(* IEC 61131-3 sources: daoli-st-library/DL_Process (part 71) *)

(* ---- FB_DL_ScrewConveyorDoseSeq.st ---- *)
(*==============================================================================
 * 组件名称 (Component)  : FB_DL_ScrewConveyorDoseSeq
 * 所属子库 (Sublibrary) : DL_Process ｜ 版本 (Version) : 1.0.0 ｜ 2026-11-24
 * 兼容性   (Platform)   : CODESYS 3.5+ / TwinCAT 3 / 汇川 InoProShop / 施耐德 Machine Expert
 *                         仅依赖 IEC 61131-3 标准库（TON / R_TRIG / ABS / MAX），零厂商私有库
 * 功能描述 (Function)   : 螺旋给料计量批次序列：预检 → 喂料（按 fFlowKgh × dt 定周期积算，
 *                         达提前量停料）→ 停料稳定 tSettle → 称量结算（算误差百分比、批次 +1、
 *                         发 bBatchDone 单拍）→ 完成相（bStart 仍 TRUE 则自动进入下一批）。
 *                         **积算口径**：dt 由定周期采样节拍 tonDt（PT = 100ms 常数）生成，
 *                         积分步长 _fDtSec = TIME_TO_LREAL(DL_SCD_DT)，且入口做 dt > EPS 闸
 *                         （防 dt ≤ 0 / 非正步长导致积分反向或除零，R4）；非采样拍不积分。
 *                         **提前量**：停料阈值 _fStopThr := fTargetKg × (1 − fTolPct/100)，
 *                         使停料后的空中料流残量落进容差带；eWeigh 再按实际 fDosedKg 结算。
 *                         **bStart = FALSE 语义（R191 二选一，本件选「降级为安全值 + 置标志」）**：
 *                         bMotorRun 落 FALSE 并回 eIdle（螺旋不得冻结保持，冻结即过量给料）。
 * 接口     (Interface)  : 输入 bEnable / bStart / bReset（上升沿）/ fTargetKg / fFlowKgh /
 *                         tSettle / tTimeout / fTolPct / bMotorFb；
 *                         输出 bMotorRun / fDosedKg / fErrPct / nBatchCnt / bBatchDone（单拍）/
 *                         eState（E_DL_ScdPhase）/ eCause（E_DL_ScdCause）/ bError / bValid。
 * 状态迁移表 (State Transition Table)：
 *   ① eIdle → ePreCheck：bEnable 且 bStart 且组态闸通过且 fTargetKg > 0 且无锁存；
 *      拍 N 进入 / 本拍行为：清 fDosedKg、fErrPct、nBatchCnt、bMotorRun=FALSE / 拍 N+1 转出。
 *   ② ePreCheck → eFeeding：预检相单拍驻留（本拍清零 fDosedKg / fErrPct，保证连续批次每批独立）；
 *      拍 N 进入 / 本拍行为：置 bMotorRun=TRUE / 拍 N+1 转出至 eFeeding。
 *   ③ eFeeding → eSettle：fDosedKg ≥ _fStopThr 或 fDosedKg ≥ fTargetKg（达量，事件优先于超时，
 *      FB51-5）；拍 N 进入 / 本拍行为：bMotorRun=FALSE、清积分节拍 / 拍 N+1 转出至 eSettle。
 *   ④ eSettle → eWeigh：tonSettle.Q（停料稳定到时）；拍 N 进入 / 本拍行为：bMotorRun=FALSE /
 *      拍 N+1 转出至 eWeigh。
 *   ⑤ eWeigh → eDone：单拍结算；本拍行为：nBatchCnt+1、置 _bBatchDoneInt（统一出口映射，
 *      FB33-1）、按 |fErrPct| 与 fTolPct 发 eBatchDone / eOutOfTol（均信息级）/ 拍 N+1 转出。
 *   ⑥ eDone → ePreCheck：bStart 仍 TRUE（连续批次）；拍 N 进入 / 本拍行为：bMotorRun=FALSE /
 *      拍 N+1 转出至 ePreCheck。⑦ eDone → eIdle：bStart 落 FALSE（前置消失，R98 两条出口）。
 *   ⑧ eFeeding → eFault：fFlowKgh < 0（eBadFlow，即时）/ 流量为 0 持续 tTimeout（eNoFlow）/
 *      总超时 tTimeout（eTimeout）/ bMotorRun 与 bMotorFb 不一致达 3s（eMotorNoFb）/
 *      全相入参非有限（eNonFinite）。锁存后由段尾迁移闸迁相（R21）。
 *   ⑨ eFault → eIdle：bReset 上升沿（R_TRIG 判 .Q）且 bEnable = FALSE（R19 穷举出口）；
 *      拍 N 进入 / 本拍行为：清锁存、成因、bMotorRun=FALSE / 拍 N+1 转出至 eIdle。
 *   ⑩ ELSE（非法枚举值）→ eFault，成因 eIllegalState（R6 兜底）。
 * 边界     (Boundary)   : ① 五个 TON 与 R_TRIG 全在 CASE 外无条件调用（R7）；tonDt / tonTotal /
 *                            tonNoFlow / tonSettle / tonMotFb 的 IN 均含 NOT .Q 自复位项（R188）。
 *                         ② 积分步长闸：_fDtSec > DL_SCD_EPS 才积分（R4 防 dt ≤ 0）；
 *                            fTargetKg ≤ EPS 时不做百分比除法，fErrPct 置 0 哨兵（除零不可达）。
 *                         ③ 浮点比较一律容差或大小比较，禁 `=`/`<>`（R4）；零流量判据为
 *                            ABS(fFlowKgh) < DL_SCD_EPS。
 *                         ④ 非有限判据：fTargetKg / fFlowKgh / fTolPct 逐拍双判（x<>x 判 NaN，
 *                            (x−x)<>0 判 Inf）。
 *                         ⑤ 无数组、无下标，故无越界风险；nBatchCnt 为 UDINT 单调累加不溢出。
 *                         ⑥ 零全局耦合（无 GVL / VAR_EXTERNAL / %I / %Q，R1 / R2）。
 * 码表     (Codes)      : 本件不占用全局数字码位（R297 零码位范式）；出口为 BOOL + ENUM，
 *                         enum E_DL_ScdPhase / E_DL_ScdCause 归属本文件（全库唯一属主，R264）。
 *                         信息级（0..9）永不置 bError；故障级（10 起）赋值处与 _bFaultLatch 三行
 *                         成对（R45），锁存回放至 bReset 沿（FB33-1）。
 * 分工声明 (Scope)      : 失重式连续给料控制（喂料闭环）归 FB_DL_ChemDosingGrav / FB_DL_BatchDosingControl；
 *                         批次报表与追溯归 DL_Process 报表件；本件只做**单批"喂料—稳定—称量"时序
 *                         与流量积算**，不做喂料闭环整定，也不做螺旋电机保护。
 * 归属     (Ownership)  : E_DL_ScdPhase / E_DL_ScdCause 归属本文件（全库唯一定义，R264）。
 * 红线自检 (Redline)    : R1 ✓ 零 GVL ｜ R2 ✓ 零 %I/%Q ｜ R3 ✓ 纯 IEC ｜ R4 ✓ dt 闸 + 除零闸 +
 *                         非有限双判 + 容差比较 ｜ R5 ✓ 逐行同行双语注释 ｜ R6 ✓ 七态 ENUM +
 *                         CASE + ELSE ｜ R7 ✓ 全部 TON/R_TRIG 在 CASE 外 ｜ R8/R9 N/A（无 METHOD）
 *                         R10 ✓ 无构造式转换（TIME_TO_LREAL / 标准函数）｜ R14 ✓ 无 PROPERTY
 *                         R15 ✓ 无保留字撞名 ｜ R17 ✓ 无数组｜ R18 ✓ bReset 用 R_TRIG 判 .Q
 *                         R19 ✓ eFault 出口 = bReset 沿 + 撤使能 ｜ R20 ✓ 稳定/供料等待相带超时
 *                         R21 ✓ 锁存与迁相分离。
 * 修订历史 (Revision)   : 2026-11-24  v1.0.0  R79-B 首版
 * 验收向量 (Acceptance) :
 *   V1 fTargetKg=10.0、fFlowKgh=3600.0（=1 kg/s）、fTolPct=1.0、tSettle=T#2S、tTimeout=T#60S：
 *      bEnable=bStart=TRUE → ePreCheck → eFeeding（bMotorRun=TRUE）；fDosedKg 每 100ms 增 0.1kg，
 *      达 9.9kg（_fStopThr）→ eSettle；2s 后 eWeigh → fErrPct≈−1.0、nBatchCnt=1、
 *      bBatchDone 单拍 TRUE（次拍 FALSE）→ eDone。
 *   V2 续 V1，bStart 保持 TRUE → eDone → ePreCheck 自动进入第 2 批；bStart 落 FALSE → 回 eIdle，
 *      nBatchCnt 清零。
 *   V3 fTargetKg=0.0 → eState=eFault、eCause=eBadConfig、bError=TRUE、bMotorRun=FALSE；
 *      bReset 上升沿且 bEnable=FALSE → 回 eIdle、bError=FALSE。
 *   V4 fFlowKgh=0.0 持续 tTimeout=T#5S → eState=eFault、eCause=eNoFlow、bError=TRUE。
 *   V5 fFlowKgh=−5.0（负流量）→ 当拍 eState=eFault、eCause=eBadFlow、bMotorRun=FALSE。
 *   V6 bMotorRun=TRUE 而 bMotorFb 保持 FALSE 超 3s → eState=eFault、eCause=eMotorNoFb。
 *============================================================================*)

(*-----------------------------------------------------------------------------
 * 枚举: E_DL_ScdPhase（螺旋给料批次相位；eFault 为安全相，仅 bReset 沿迁出）
 *----------------------------------------------------------------------------*)
TYPE E_DL_ScdPhase :
(
    eIdle     := 0,    // 空闲：电机停，计数值清零 / Idle: motor stopped, counters cleared
    ePreCheck := 10,   // 预检相：单拍，置电机启动命令 / Pre-check: single scan, arm the motor command
    eFeeding  := 20,   // 喂料相：电机运行，按流量 × dt 积算 / Feeding: motor on, integrate flow times dt
    eSettle   := 30,   // 稳定相：停料后等空中料流落净 / Settle: motor off, waiting for the in-flight material
    eWeigh    := 40,   // 称量相：单拍结算误差与批次 / Weigh: single-scan settlement of error and batch count
    eDone     := 50,   // 完成相：本批完成，等下一批或退出 / Done: batch finished, waiting for the next one
    eFault    := 90    // 故障安全相：锁存成因，电机全停 / Fault safe phase: latched cause, motor stopped
);
END_TYPE

(*-----------------------------------------------------------------------------
 * 枚举: E_DL_ScdCause（成因码；信息级 = 0..9，故障级 = 10 起）
 *----------------------------------------------------------------------------*)
TYPE E_DL_ScdCause :
(
    eNone       := 0,   // 信息级：无事件 / Info: no event
    eBatchDone  := 1,   // 信息级：一批完成且误差在容差内 / Info: batch completed within tolerance
    eOutOfTol   := 2,   // 信息级：一批完成但误差超容差（记录，不锁存）/ Info: batch completed out of tolerance, recorded only
    eSettling   := 3,   // 信息级：进入停料稳定相 / Info: entering the settle phase
    eBadConfig  := 10,  // 故障级：目标重量 / 容差 / 时间参数越域 / Fault: target, tolerance or time parameter out of domain
    eNonFinite  := 11,  // 故障级：入参非有限 / Fault: non-finite input
    eBadFlow    := 12,  // 故障级：流量为负 / Fault: negative flow
    eNoFlow     := 13,  // 故障级：流量为零持续超时（供料中断）/ Fault: zero flow persisted beyond the timeout
    eTimeout    := 14,  // 故障级：喂料总超时 / Fault: total feeding timeout
    eMotorNoFb  := 15,  // 故障级：电机命令与反馈不一致超 3s / Fault: motor command and feedback mismatch beyond 3 s
    eIllegalState := 16 // 故障级：非法状态枚举值 / Fault: illegal state enum value
);
END_TYPE

FUNCTION_BLOCK FB_DL_ScrewConveyorDoseSeq
VAR_INPUT
    bEnable    : BOOL := FALSE;        // 使能：FALSE 停电机并回 eIdle / Enable, FALSE stops the motor and returns to idle
    bStart     : BOOL := FALSE;        // 启动（电平）：FALSE 本批中止并回 eIdle / Start level, FALSE aborts the batch
    bReset     : BOOL := FALSE;        // 复位（上升沿，需同时 bEnable=FALSE）/ Reset rising edge, requires bEnable FALSE
    fTargetKg  : LREAL := 0.0;         // 批次目标重量，域 > 0 [kg] / Batch target weight, domain > 0
    fFlowKgh   : LREAL := 0.0;         // 当前给料流量（瞬时，来自流量计）[kg/h] / Instantaneous feed flow from the flow meter
    tSettle    : TIME := T#2S;         // 停料后稳定延时，域 0..1h [s] / Settle delay after the motor stops, domain 0..1h
    tTimeout   : TIME := T#60S;        // 喂料总超时，域 ≥ 100ms [s] / Total feeding timeout, domain >= 100ms
    fTolPct    : LREAL := 1.0;         // 允许误差，域 (0,100) [%] / Allowed error in percent, domain (0,100)
    bMotorFb   : BOOL := FALSE;        // 螺旋电机运行反馈（TRUE = 在转）[-] / Screw motor running feedback
END_VAR
VAR_OUTPUT
    bMotorRun  : BOOL;                 // 螺旋电机启动命令（电平）[-] / Screw motor run command, level
    fDosedKg   : LREAL := 0.0;         // 本批累计给料量 [kg] / Accumulated dose of this batch
    fErrPct    : LREAL := 0.0;         // 本批误差百分比（正 = 超量）[%] / Batch error percentage, positive means over-dose
    nBatchCnt  : UDINT := 0;           // 已完成批次数 [批] / Completed batch counter
    bBatchDone : BOOL;                 // 批次完成单拍脉冲（段 1 预置，统一出口映射）[-] / Single-scan batch-done pulse
    eState     : E_DL_ScdPhase;        // 状态出口（段尾单点映射）[-] / State outlet mapped at the tail
    eCause     : E_DL_ScdCause;        // 成因码出口（故障期锁存回放）[-] / Cause code outlet
    bError     : BOOL;                 // 故障锁存标志 [-] / Fault latch flag
    bValid     : BOOL;                 // 序列有效回执（喂料/稳定相且无锁存）[-] / Sequence validity receipt
END_VAR
VAR
    _eState      : E_DL_ScdPhase := E_DL_ScdPhase.eIdle;   // 内部相位（CASE 唯一写入目标）[-] / Internal phase
    _bFaultLatch : BOOL := FALSE;                          // 故障锁存位（仅 bReset 沿清除）[-] / Fault latch bit
    _eCauseLatch : E_DL_ScdCause := E_DL_ScdCause.eNone;    // 锁存成因码（FB33-1 锁存回放）[-] / Latched cause code
    _eCauseTmp   : E_DL_ScdCause := E_DL_ScdCause.eNone;    // 本拍首因中间量（段 8 组态闸用）[-] / First cause of this scan
    _bCfgOk      : BOOL := TRUE;                           // 组态与入参闸通过标志 [-] / Configuration gate flag
    _bResetPulse : BOOL := FALSE;                          // bReset 上升沿快照（R18）[-] / bReset rising-edge snapshot
    _bBatchDoneInt : BOOL := FALSE;                        // 批次完成内部单拍位（统一出口映射）[-] / Internal single-scan batch-done bit
    _fDtSec      : LREAL := 0.0;                           // 积分步长：[s] / Integration step in seconds
    _bDtOk       : BOOL := FALSE;                          // 积分步长有效性（dt > EPS）[-] / Integration step validity
    _fStopThr    : LREAL := 0.0;                           // 停料阈值 = 目标 × (1 − 容差%) [kg] / Stop threshold of the feed
    _fStepKg     : LREAL := 0.0;                           // 本采样拍积算增量 [kg] / Dose increment of this sampling scan
    _fErrCalc    : LREAL := 0.0;                           // 误差百分比中间量 [%] / Error percentage intermediate
    _bMotMismatch : BOOL := FALSE;                         // 电机命令与反馈不一致标志 [-] / Motor command and feedback mismatch
    _bMotRunPrev  : BOOL := FALSE;                         // 上一拍电机命令快照（段 4 不一致判据用，一拍延迟）/ Motor command snapshot of the last scan
    rtReset      : R_TRIG;                                 // bReset 边沿实例（段 4 无条件调用，R18）/ bReset edge instance called unconditionally
    tonDt        : TON;                                    // 定周期采样节拍（段 4 无条件调用）/ Fixed-period sampling tick
    tonTotal     : TON;                                    // 喂料总超时（段 4 无条件调用）/ Total feeding timeout
    tonNoFlow    : TON;                                    // 零流量持续判（段 4 无条件调用）/ Zero-flow persistence timer
    tonSettle    : TON;                                    // 停料稳定延时（段 4 无条件调用）/ Settle delay timer
    tonMotFb     : TON;                                    // 电机反馈不一致持续判（段 4 无条件调用）/ Motor feedback mismatch timer
END_VAR
VAR CONSTANT
    DL_SCD_ZERO      : LREAL := 0.0;            // 浮点零基准 [-] / Float zero base
    DL_SCD_ONE       : LREAL := 1.0;            // 浮点一基准 [-] / Float one base
    DL_SCD_HUNDRED   : LREAL := 100.0;          // 百分比基数 [%] / Percent base
    DL_SCD_SEC_HOUR  : LREAL := 3600.0;         // 每小时秒数（kg/h → kg）[s/h] / Seconds per hour converting kg/h to kg
    DL_SCD_EPS       : LREAL := 1.0E-6;         // 浮点同值/正步长容差 [-] / Float equality and positive-step tolerance
    DL_SCD_DT        : TIME := T#100MS;         // 采样节拍（积分步长来源）[s] / Sampling tick, the integration step source
    DL_SCD_FB_WIN    : TIME := T#3S;            // 电机反馈不一致持续窗 [s] / Motor feedback mismatch window
    DL_SCD_T_MIN     : TIME := T#100MS;         // 超时参数下限 [s] / Lower bound of the timeout parameters
    DL_SCD_T_MAX     : TIME := T#1H;            // 稳定/超时参数上限 [s] / Upper bound of the settle and timeout parameters
    DL_SCD_BATCH_INC : UDINT := 1;              // 批次计数步长（UDINT 显式常量）[批] / Batch counter increment
END_VAR

(* —— 段 1：单拍位与动作出口预置（不清锁存 / 累加量，FB32-1） —— *)
bBatchDone     := FALSE;                               // 单拍批次沿每拍预清 / Single-scan batch edge preset FALSE every scan
bMotorRun      := FALSE;                               // 电机命令预置（安全侧：默认不动作）/ Motor command preset, safe side
_bBatchDoneInt := FALSE;                               // 内部单拍位预清 / Internal single-scan bit preset
_bCfgOk        := TRUE;                                // 组态闸标志复位 / Configuration flag reset
_eCauseTmp     := E_DL_ScdCause.eNone;                  // 当拍首因复位 / Scan cause reset

(* —— 段 2：步长与阈值换算（浮点域闸前置） —— *)
_fDtSec   := TIME_TO_LREAL(DL_SCD_DT);                 // 采样节拍换算为秒（标准转换，R10）/ Sampling tick converted to seconds
IF _fDtSec > DL_SCD_EPS THEN
    _bDtOk := TRUE;                                    // 步长为正：允许积分 / Positive step: integration allowed
ELSE
    _bDtOk := FALSE;                                   // 步长非正：拒绝积分（R4 防 dt <= 0）/ Non-positive step: integration refused
END_IF
_fStopThr := DL_SCD_ZERO;                              // 停料阈值预置零 / Stop threshold preset
_fErrCalc := DL_SCD_ZERO;                               // 误差中间量预置零 / Error intermediate preset

(* —— 段 3：组态与入参域闸（R272 全量枚举浮点与时间引脚） —— *)
IF (fTargetKg <> fTargetKg) OR ((fTargetKg - fTargetKg) <> DL_SCD_ZERO)
    OR (fFlowKgh <> fFlowKgh) OR ((fFlowKgh - fFlowKgh) <> DL_SCD_ZERO)
    OR (fTolPct <> fTolPct) OR ((fTolPct - fTolPct) <> DL_SCD_ZERO) THEN
    _bCfgOk    := FALSE;                               // 入参非有限 / Non-finite input
    _eCauseTmp := E_DL_ScdCause.eNonFinite;            // 故障级：非有限入参 / Fault: non-finite input
END_IF
IF _bCfgOk THEN
    IF fTargetKg <= DL_SCD_EPS THEN
        _bCfgOk    := FALSE;                           // 目标重量非正 / Target weight not positive
        _eCauseTmp := E_DL_ScdCause.eBadConfig;        // 故障级：组态非法 / Fault: bad configuration
    ELSIF (fTolPct <= DL_SCD_EPS) OR (fTolPct >= DL_SCD_HUNDRED) THEN
        _bCfgOk    := FALSE;                           // 容差越域（0,100）/ Tolerance out of domain
        _eCauseTmp := E_DL_ScdCause.eBadConfig;        // 故障级：组态非法 / Fault: bad configuration
    ELSIF (tTimeout < DL_SCD_T_MIN) OR (tTimeout > DL_SCD_T_MAX) THEN
        _bCfgOk    := FALSE;                           // 超时参数越域 / Timeout out of domain
        _eCauseTmp := E_DL_ScdCause.eBadConfig;        // 故障级：组态非法 / Fault: bad configuration
    ELSIF tSettle > DL_SCD_T_MAX THEN
        _bCfgOk    := FALSE;                           // 稳定延时越上限 / Settle delay above the upper bound
        _eCauseTmp := E_DL_ScdCause.eBadConfig;        // 故障级：组态非法 / Fault: bad configuration
    ELSIF fFlowKgh < DL_SCD_ZERO THEN
        _bCfgOk    := FALSE;                           // 流量为负（传感器或工艺异常）/ Negative flow from the meter or process
        _eCauseTmp := E_DL_ScdCause.eBadFlow;          // 故障级：负流量 / Fault: negative flow
    END_IF
END_IF
IF _bCfgOk THEN
    (* 停料阈值 = 目标 × (1 − 容差%/100)；除数 100 为常量，除零结构性不可达 *)
    _fStopThr := fTargetKg * (DL_SCD_ONE - (fTolPct / DL_SCD_HUNDRED));
    IF _fStopThr <= DL_SCD_ZERO THEN
        _fStopThr := DL_SCD_ZERO;                      // 阈值负值兜底归零 / Clamp a negative threshold to zero
    END_IF
END_IF

(* —— 段 4：边沿与定时器（CASE 外无条件调用，R7；IN 均含 NOT .Q 自复位，R188） —— *)
rtReset(CLK := bReset);                                // bReset 边沿无条件刷新（R18）/ bReset edge refreshed unconditionally
_bResetPulse := rtReset.Q;                             // 边沿快照 / Edge snapshot
tonDt(IN := (_eState = E_DL_ScdPhase.eFeeding) AND (NOT tonDt.Q) AND (NOT _bFaultLatch),
      PT := DL_SCD_DT);                                // 喂料相定周期积分节拍 / Fixed-period integration tick while feeding
tonTotal(IN := (_eState = E_DL_ScdPhase.eFeeding) AND (NOT tonTotal.Q) AND (NOT _bFaultLatch),
         PT := tTimeout);                              // 喂料总超时 / Total feeding timeout
tonNoFlow(IN := (_eState = E_DL_ScdPhase.eFeeding) AND (ABS(fFlowKgh) < DL_SCD_EPS)
               AND (NOT tonNoFlow.Q) AND (NOT _bFaultLatch),
          PT := tTimeout);                             // 零流量持续判（供料中断）/ Zero-flow persistence check
tonSettle(IN := (_eState = E_DL_ScdPhase.eSettle) AND (NOT tonSettle.Q) AND (NOT _bFaultLatch),
          PT := tSettle);                              // 停料稳定延时 / Settle delay
_bMotMismatch := (_bMotRunPrev AND (NOT bMotorFb)) OR ((NOT _bMotRunPrev) AND bMotorFb);   // 命令与反馈不一致（用上一拍命令快照）/ Command and feedback mismatch using the last-scan command
tonMotFb(IN := _bMotMismatch AND (_eState = E_DL_ScdPhase.eFeeding)
              AND (NOT tonMotFb.Q) AND (NOT _bFaultLatch),
         PT := DL_SCD_FB_WIN);                         // 仅喂料相监视反馈一致性 / Feedback consistency monitored while feeding only

(* —— 段 5：误差百分比刷新（除零闸：目标重量非正时置零哨兵，R4） —— *)
IF fTargetKg > DL_SCD_EPS THEN
    _fErrCalc := ((fDosedKg - fTargetKg) / fTargetKg) * DL_SCD_HUNDRED;   // 误差百分比 / Error percentage
    fErrPct   := _fErrCalc;                                               // 误差出口 / Error outlet
ELSE
    fErrPct := DL_SCD_ZERO;                                               // 目标非正：置零哨兵（除零不可达）/ Zero sentinel, division unreachable
END_IF

(* —— 段 6：状态机主体（唯一相位写入点；故障只置锁存，迁相由段 8 统一执行） —— *)
CASE _eState OF
    E_DL_ScdPhase.eIdle :
        bMotorRun := FALSE;                            // 空闲：电机不动作 / Idle: motor idle
        fDosedKg  := DL_SCD_ZERO;                      // 累计量清零 / Dose counter cleared
        fErrPct   := DL_SCD_ZERO;                      // 误差清零 / Error cleared
        nBatchCnt := 0;                                // 批次计数清零 / Batch counter cleared
        IF bEnable AND bStart AND _bCfgOk AND (fTargetKg > DL_SCD_EPS) AND (NOT _bFaultLatch) THEN
            eCause  := E_DL_ScdCause.eNone;            // 信息级：无事件 / Info: no event
            _eState := E_DL_ScdPhase.ePreCheck;        // 迁移①：进入预检相 / Move to pre-check
        END_IF

    E_DL_ScdPhase.ePreCheck :
        IF (NOT bEnable) OR (NOT bStart) THEN
            bMotorRun := FALSE;                        // 失能：电机停 / Disabled: motor stopped
            eCause    := E_DL_ScdCause.eNone;          // 信息级：无事件 / Info: no event
            _eState   := E_DL_ScdPhase.eIdle;          // 回空闲相 / Back to idle
        ELSE
            fDosedKg  := DL_SCD_ZERO;                  // 每批起点：累计量清零 / Batch start: dose counter cleared
            fErrPct   := DL_SCD_ZERO;                  // 每批起点：误差清零 / Batch start: error cleared
            bMotorRun := TRUE;                         // 迁移②：预检通过，启动螺旋 / Pre-check passed: start the screw
            eCause    := E_DL_ScdCause.eNone;          // 信息级：无事件 / Info: no event
            _eState   := E_DL_ScdPhase.eFeeding;       // 进入喂料相 / Move to feeding
        END_IF

    E_DL_ScdPhase.eFeeding :
        bMotorRun := TRUE;                             // 喂料相电机保持运行 / Motor stays on while feeding
        IF (NOT bEnable) OR (NOT bStart) THEN
            bMotorRun := FALSE;                        // 失能：电机停 / Disabled: motor stopped
            eCause    := E_DL_ScdCause.eNone;          // 信息级：无事件 / Info: no event
            _eState   := E_DL_ScdPhase.eIdle;          // 回空闲相 / Back to idle
        ELSE
            (* 定周期积算：只有节拍拍且步长为正才积分（R4） *)
            IF tonDt.Q AND _bDtOk THEN
                _fStepKg  := (fFlowKgh * _fDtSec) / DL_SCD_SEC_HOUR;   // 增量 = 流量 × dt / 3600 [kg]
                fDosedKg  := fDosedKg + _fStepKg;                      // 累计给料量 / Accumulate the dose
            END_IF
            IF fFlowKgh < DL_SCD_ZERO THEN
                IF NOT _bFaultLatch THEN
                    _eCauseLatch := E_DL_ScdCause.eBadFlow;            // 故障级：负流量 / Fault: negative flow
                    _bFaultLatch := TRUE;                              // 置故障锁存（迁相由段 8，R21）/ Latch the fault
                END_IF
            ELSIF tonNoFlow.Q THEN
                IF NOT _bFaultLatch THEN
                    _eCauseLatch := E_DL_ScdCause.eNoFlow;             // 故障级：供料中断 / Fault: feed interrupted
                    _bFaultLatch := TRUE;                              // 置故障锁存 / Latch the fault
                END_IF
            ELSIF tonTotal.Q THEN
                IF NOT _bFaultLatch THEN
                    _eCauseLatch := E_DL_ScdCause.eTimeout;            // 故障级：喂料总超时 / Fault: total feeding timeout
                    _bFaultLatch := TRUE;                              // 置故障锁存 / Latch the fault
                END_IF
            ELSIF tonMotFb.Q THEN
                IF NOT _bFaultLatch THEN
                    _eCauseLatch := E_DL_ScdCause.eMotorNoFb;          // 故障级：电机反馈不一致 / Fault: motor feedback mismatch
                    _bFaultLatch := TRUE;                              // 置故障锁存 / Latch the fault
                END_IF
            ELSIF (fDosedKg >= _fStopThr) OR (fDosedKg >= fTargetKg) THEN
                bMotorRun := FALSE;                                    // 迁移③：达提前量，停料 / Reached the threshold: stop the feed
                eCause    := E_DL_ScdCause.eSettling;                  // 信息级：进入稳定相 / Info: entering settle
                _eState   := E_DL_ScdPhase.eSettle;                    // 进入稳定相 / Move to settle
            END_IF
        END_IF

    E_DL_ScdPhase.eSettle :
        bMotorRun := FALSE;                            // 稳定相电机保持停止 / Motor stays off while settling
        IF (NOT bEnable) OR (NOT bStart) THEN
            eCause  := E_DL_ScdCause.eNone;            // 信息级：无事件 / Info: no event
            _eState := E_DL_ScdPhase.eIdle;            // 回空闲相 / Back to idle
        ELSIF tonSettle.Q THEN
            eCause  := E_DL_ScdCause.eNone;            // 信息级：无事件 / Info: no event
            _eState := E_DL_ScdPhase.eWeigh;           // 迁移④：稳定到时进入称量相 / Settle elapsed: move to weigh
        END_IF

    E_DL_ScdPhase.eWeigh :
        bMotorRun      := FALSE;                       // 称量相电机停止 / Motor off during settlement
        nBatchCnt      := nBatchCnt + DL_SCD_BATCH_INC; // 迁移⑤：批次计数 +1 / Increment the batch counter
        _bBatchDoneInt := TRUE;                        // 批次完成内部单拍位置位 / Internal single-scan batch bit
        IF ABS(fErrPct) > fTolPct THEN
            eCause := E_DL_ScdCause.eOutOfTol;         // 信息级：误差超容差（记录，不锁存）/ Info: out of tolerance, recorded only
        ELSE
            eCause := E_DL_ScdCause.eBatchDone;        // 信息级：批次合格完成 / Info: batch completed within tolerance
        END_IF
        _eState := E_DL_ScdPhase.eDone;                // 进入完成相 / Move to done

    E_DL_ScdPhase.eDone :
        bMotorRun := FALSE;                            // 完成相电机停止 / Motor off in the done phase
        IF NOT bStart THEN
            eCause  := E_DL_ScdCause.eNone;            // 信息级：无事件 / Info: no event
            _eState := E_DL_ScdPhase.eIdle;            // 迁移⑦：前置消失回空闲 / Start gone: back to idle
        ELSIF NOT bEnable THEN
            eCause  := E_DL_ScdCause.eNone;            // 信息级：无事件 / Info: no event
            _eState := E_DL_ScdPhase.eIdle;            // 失能回空闲 / Disabled: back to idle
        ELSIF bStart AND bEnable THEN
            eCause  := E_DL_ScdCause.eNone;            // 信息级：无事件 / Info: no event
            _eState := E_DL_ScdPhase.ePreCheck;        // 迁移⑥：连续批次 / Continuous batches
        END_IF

    E_DL_ScdPhase.eFault :
        bMotorRun := FALSE;                            // 故障相：电机全停（安全侧）/ Fault phase: motor stopped
        IF _bResetPulse AND (NOT bEnable) THEN
            _bFaultLatch := FALSE;                     // 迁移⑨：清故障锁存 / Clear the fault latch
            _eCauseLatch := E_DL_ScdCause.eNone;       // 清锁存成因 / Clear the latched cause
            eCause       := E_DL_ScdCause.eNone;       // 出口同步归零 / Outlet follows
            fDosedKg     := DL_SCD_ZERO;               // 累计量清零 / Dose counter cleared
            fErrPct      := DL_SCD_ZERO;               // 误差清零 / Error cleared
            _eState      := E_DL_ScdPhase.eIdle;       // 回空闲相 / Back to idle
        END_IF

ELSE
    (* 迁移⑩：非法枚举兜底（R6） *)
    IF NOT _bFaultLatch THEN
        _eCauseLatch := E_DL_ScdCause.eIllegalState;   // 故障级：非法状态 / Fault: illegal state
        _bFaultLatch := TRUE;                          // 置故障锁存 / Latch the fault
    END_IF
END_CASE

(* —— 段 7：组态闸失败处理（锁存与迁相分离，R21） —— *)
IF (NOT _bCfgOk) AND (NOT _bFaultLatch) THEN
    _eCauseLatch := _eCauseTmp;                        // 锁存首因（组态闸）/ Latch the configuration cause
    _bFaultLatch := TRUE;                              // 置故障锁存 / Latch the fault
END_IF

(* —— 段 8：段尾故障迁移闸 + 故障相动作全撤（FB50-1④） —— *)
IF _bFaultLatch AND (_eState <> E_DL_ScdPhase.eFault) THEN
    _eState := E_DL_ScdPhase.eFault;                   // 锁存即迁相 / Latch forces the fault phase
END_IF
IF _eState = E_DL_ScdPhase.eFault THEN
    bMotorRun := FALSE;                                // 故障相动作全撤（含同拍迁入）/ Motor withdrawn in fault
END_IF

(* —— 段 9：统一出口（状态映射 + 单拍位映射 + 锁存回放） —— *)
eState     := _eState;                                 // 相位映射 / Phase mapping
bBatchDone := _bBatchDoneInt;                          // 单拍批次沿统一映射（FB33-1 两段式）/ Single-scan batch edge mapped here
bError     := _bFaultLatch;                            // 故障标志取锁存位 / Fault flag from the latch
IF _bFaultLatch THEN
    eCause := _eCauseLatch;                            // 故障期回放锁存码（FB33-1）/ Replay the latched code
END_IF
bValid := ((_eState = E_DL_ScdPhase.eFeeding) OR (_eState = E_DL_ScdPhase.eSettle))
          AND (NOT _bFaultLatch);                      // 喂料/稳定相且无锁存时有效 / Valid while feeding or settling without a latch
_bMotRunPrev := bMotorRun;                             // 电机命令快照更新（唯一写入点，段 4 用）/ Motor command snapshot, single write point
END_FUNCTION_BLOCK

(* ---- FB_DL_SipLineSterilSeq.st ---- *)
(*
    FB_DL_SipLineSterilSeq —— 管路 SIP 蒸汽灭菌顺控（排凝 → 升温 → 保温窗 → 冷却 → 放行）
    ------------------------------------------------------------------
    组件名称  : FB_DL_SipLineSterilSeq
    分类      : DL_Process / Sterilization
    前缀      : FB_DL_
    版本      : 1.0.0
    溯源      : 借鉴组织 —— T2-2 LBP 基础工艺（矩阵行 163）：仅借鉴
                「命令 → 监视 → 判定」三段分层骨架的公开语义；次源 T2-8
                ISA-88 相语义公开条款（相 / 状态命名惯例）；clean-room
                声明 —— 保温窗断点重计与温度判据 100% 自有，零代码行复制；
                SIP 121 ℃ 最低承诺属公开工程惯例条款（下界 100 ℃ 为本件
                组态锁存闸，可调）。
    平台      : 纯 IEC 61131-3（ENUM + CASE + TON / R_TRIG + TIME 算术），
                CODESYS 3.5 / TwinCAT 3 / InoProShop / Machine Expert 通用
    作者      : 道莅代码库 · PLC编程专家（R72 构建轮 · 批 4 · 序号 12）
    ------------------------------------------------------------------
    功能说明  : 管路蒸汽 SIP（Sterilize-In-Place）连续工艺段顺控：
                eIdle →（bEn ∧ 组态闸）eDrain（排凝，bDrainDone 反馈或
                tDrainTimeout 超时）→ eHeatUp（开蒸汽升温，fTempC 达
                fHoldTempSet 迁入）→ eHold（保温窗 TON 计时）→ eCooldown
                （关蒸汽，温度回落确认）→ eDone（bSterilized 放行保持）→
                eIdle（批界）。
                安全核心口径：
                ① fTempC 非有限（探头断线）→ **故障锁存 + 双输出立即关断**
                   ——温度状态不明不得放行，宁可重灭菌；
                ② 保温窗断点重计（SIP 无菌保证不容断点续计）：eHold 相内
                   fTempC 跌破 fHoldTempSet（每拍取本拍实时值，R42 本拍
                   复验口径）→ 计时中止回 eHeatUp + 扰动计数 +1，恢复后
                   TON 从零重计——断点续计等于伪造无菌时长，写死禁用；
                ③ fHoldTempSet 越承诺段（< 100 ℃）→ 组态锁存（SIP 公开
                   最低承诺 121 ℃ 工程惯例，下界闸定 100 ℃ 并留调参会空间
                   ——承诺下界以常量声明，单探头承诺段声明见边界八）；
                ④ 失能 → 双输出（bDrainCmd / bSteamCmd）清零 + bSterilized
                   撤销 + 状态回 eIdle（停机相输出清零，R57）；故障锁存保留，
                   复位沿解除；
                ⑤ 迁入 eHold 相与每拍判温均取本拍实时值（迁入拍即计时使能，
                   无跨拍陈旧判据）。
                冷却放行口径：eCooldown 以 fTempC < fHoldTempSet 确认回落
                （防高温放行烫尾），回落即 eDone；bSterilized 为**保持型**
                放行位（批界 = bEn 撤除或复位沿时清除）。
    错误码    : 16#0005_0640 工艺温度非有限（探头断线 / ADC 故障），双输出
                            立即关断，锁存至复位沿 —— 故障级
                16#0005_0641 排凝超时（eDrain 驻留超 tDrainTimeout），锁存
                            至复位沿 —— 故障级
                16#0005_0642 保温设定越承诺段（fHoldTempSet < 100 ℃ 或非
                            有限），锁存至复位沿 —— 故障级
                16#0005_0643 保温窗 / 排凝超时组态非正（tHoldTime /
                            tDrainTimeout <= 0），锁存至复位沿 —— 故障级
                加码反证句（R90）：0640 由「双输出关断 + eHealth 语义温度
                断线」唯一观测；0641 / 0642 / 0643 成因互斥且调用方可自证
                （反馈时序 / 组态表），输出组合（同为 eFault + bError）不可
                互换还原成因，维修动作各异，故各立一码；保温跌破扰动以
                uDisturbCount 专位观测（R90 不加码：扰动事件已有独立可观
                测出口，不重复发码）。
    码位总账  : 16#0005_0640 用 ｜ 16#0005_0641 用 ｜ 16#0005_0642 用 ｜
                16#0005_0643 用
                （0630 / 0631 已由 FB_DL_RejectBlowCtrl 占用，本件不占）
    边界与披露: 一 双 TON（tonDrain / tonHold）与 R_TRIG（rtReset）每拍
                   **无条件调用**（规则 ⑦），IN 为显式条件变量（R145 相驻留
                   口径：tonDrain IN = 排凝相驻留，tonHold IN = 保温相驻留
                   ∧ 本拍温度达标）；
                二 零全局变量、零 VAR_EXTERNAL、零物理地址；
                三 归属 Ownership：E_DL_SipPhase 属主为本文件（全库唯一定义，
                   R264），引用件只引用不重声明；
                四 状态机 ENUM + CASE 必带 ELSE 兜底（非法枚举值 → eFault
                   锁存）+ 段 5b 统一故障迁入闸（R274 迁入完备性）；
                五 域闸逐项点名（R272）：fTempC（非有限闸）+ fHoldTempSet
                   （非有限与承诺段闸）全部浮点引脚入闸；
                六 时间量纲口径：tHoldTime / tDrainTimeout 均为 TIME 引脚
                   （内部毫秒），保温剩余 uHoldRemain 以秒发布（TIME_TO_DINT
                   毫秒差 ÷ 常量除子 1000，零除法面，R382 常量除子级联）；
                七 单探头承诺段声明：本件按单工艺温度探头承诺（多点冷点
                   归上位编排，数组版不立防拆件凑数）；fHoldTempSet 默认
                   121.0 ℃ 仅为 SIP 工程惯例参考值，非承诺；
                八 分工声明：FB_DL_CipCleaningSeq（化学清洗顺控）、
                   FB_DL_AutoclaveSterilSeq（灭菌釜批次）、
                   FB_DL_TunnelPasteurizerSeq（隧道巴氏）——本件专管
                   **管路蒸汽 SIP 连续工艺段**，互引不互代；
                九 复位沿作用域（R311）：清全部锁存 + 清锁存码 + 迁 eIdle +
                   清 bSterilized（批界复位）+ 清扰动计数（批次台账随批清），
                   **不清**自动统计类（本件无）；
                十 依赖声明：仅 Standard.library（TON / R_TRIG），零厂商
                   方言。
    验收向量  : V1 正常批次：排凝反馈 → 升温达标 → 保温 tHoldTime → 冷却
                回落 → bSterilized 保持，uDisturbCount = 0；
                V2 保温中跌破设定 → 回 eHeatUp + uDisturbCount + 1，恢复后
                保温从零重计（断点重计口径自证）；
                V3 fTempC = NaN → 0640 锁存 + 双输出关断；
                V4 fHoldTempSet = 90 ℃ → 0642 锁存；V5 tHoldTime = T#0S →
                0643 锁存；V6 排凝超时 → 0641 锁存；V7 失能 → 双输出清零 +
                bSterilized 撤销；V8 复位沿 → 解锁回 eIdle。
                算法已证（脚本）：未跑 ｜ 编译器已证（三平台）：未跑
    修订记录  : 2026-11-23 v1.0.0 首次入库（R72 构建轮 · 批 4 · 序号 12）
*)
TYPE E_DL_SipPhase :
(
    eIdle     := 0,                        // 空闲：等使能与组态闸 / idle, waiting for the enable
    eDrain    := 10,                       // 排凝：等反馈或超时 / drain, waiting for the feedback
    eHeatUp   := 20,                       // 升温：开蒸汽等达标 / heat up, the steam on
    eHold     := 30,                       // 保温窗：TON 计时，跌破重计 / hold, the timed window
    eCooldown := 40,                       // 冷却：关蒸汽等回落 / cooldown, the steam off
    eDone     := 50,                       // 放行：bSterilized 保持相 / done, the release phase
    eFault    := 60                        // 故障：锁存待复位 / fault, latched until the reset
);
END_TYPE

FUNCTION_BLOCK FB_DL_SipLineSterilSeq
VAR_INPUT
    fTempC        : LREAL;                 (* 工艺温度探头（单探头承诺段），[摄氏度]，非有限即探头故障 / the process temperature in degC *)
    bDrainDone    : BOOL := FALSE;         (* 排凝完成反馈，[标志]，引脚注入 / the drain done feedback *)
    fHoldTempSet  : LREAL := 121.0;        (* 保温承诺温度，[摄氏度]，禁 < 100 / 非有限（默认 121 为 SIP 惯例参考值）/ the hold temperature setpoint *)
    tHoldTime     : TIME := T#1800S;       (* 保温窗，[ms]，禁非正 / the hold window duration *)
    tDrainTimeout : TIME := T#300S;        (* 排凝超时，[ms]，禁非正 / the drain timeout *)
    bEn           : BOOL := FALSE;         (* 使能，[标志]，FALSE 双输出清零回 eIdle（锁存保留）/ the enable *)
    bReset        : BOOL := FALSE;         (* 故障复位，[标志]，上升沿唯一解除 / the fault reset *)
END_VAR
VAR_OUTPUT
    bDrainCmd   : BOOL := FALSE;           (* 排凝指令出口，[标志]，故障 / 失能为 FALSE / the drain command outlet *)
    bSteamCmd   : BOOL := FALSE;           (* 蒸汽指令出口，[标志]，故障 / 失能为 FALSE（安全侧关断）/ the steam command outlet *)
    bSterilized : BOOL := FALSE;           (* 灭菌放行出口（保持型，批界清除）[标志] / the sterilized release outlet *)
    uHoldRemain : UDINT := 0;              (* 保温剩余倒计时（HMI），[秒]，非保温相为 0 / the hold remaining seconds *)
    uDisturbCount: UDINT := 0;             (* 保温跌破扰动计数（批界复位）[次] / the hold disturbance count *)
    eState      : E_DL_SipPhase := E_DL_SipPhase.eIdle; // 主状态机当前态 [状态] / the current state
    bError      : BOOL := FALSE;           (* 故障标志，与锁存同源（R191）/ the fault flag from the latch *)
    nErrCode    : UDINT := 16#0000_0000;   (* 错误码，0 = 正常，故障锁存回放（R187）/ the error id *)
END_VAR
VAR
    _bInit      : BOOL := FALSE;           (* 首拍初始化标志（R310）/ the first scan flag *)
    _eState     : E_DL_SipPhase := E_DL_SipPhase.eIdle; // 内部状态寄存器 / the internal state register
    _bFault     : BOOL := FALSE;           (* 故障锁存副本，仅复位沿解除 / the fault latch copy *)
    _nCodeLatch : UDINT := 0;              (* 锁存成因码，故障期回放 / the latched cause code *)
    _bCfgBad    : BOOL := FALSE;           (* 组态非法标志（逐拍重算，仅用于首次锁存）/ the config fault flag *)
    _bTInBad    : BOOL := FALSE;           (* 温度非有限标志（逐拍重算，R272 闸）/ the temperature invalid flag *)
    _bTempOk    : BOOL := FALSE;           (* 本拍温度达标实时判据（R42 本拍复验）/ the live temperature verdict *)
    _bDrain     : BOOL := FALSE;           (* 排凝指令内部位（统一出口映射）/ the internal drain bit *)
    _bSteam     : BOOL := FALSE;           (* 蒸汽指令内部位（统一出口映射）/ the internal steam bit *)
    _bReleased  : BOOL := FALSE;           (* 放行内部锁存（eDone 相保持）/ the internal release latch *)
    nRemainMs   : DINT := 0;               (* 保温剩余毫秒中间量 [ms] / the remaining milliseconds temporary *)
    rtReset     : R_TRIG;                  (* 复位沿实例（无条件调用）/ the reset edge instance *)
    tonDrain    : TON;                     (* 排凝超时看门狗（无条件调用）/ the drain watchdog timer *)
    tonHold     : TON;                     (* 保温窗计时（无条件调用）/ the hold window timer *)
END_VAR
VAR CONSTANT
    DL_SIP_CODE_TEMP : UDINT := 16#0005_0640; // 温度非有限故障码 [码] / the probe fault code
    DL_SIP_CODE_DRAIN: UDINT := 16#0005_0641; // 排凝超时故障码 [码] / the drain timeout code
    DL_SIP_CODE_SET  : UDINT := 16#0005_0642; // 保温设定越承诺段故障码 [码] / the setpoint fault code
    DL_SIP_CODE_TIME : UDINT := 16#0005_0643; // 时间组态非正故障码 [码] / the time config fault code
    DL_SIP_TSETMIN   : LREAL := 100.0;       (* 保温承诺温度下界（SIP 公开最低承诺 121 ℃，下界闸 100 ℃ 可调参会）[摄氏度] / the setpoint promise lower bound *)
    DL_SIP_TZERO     : LREAL := 0.0;         (* 浮点零哨兵 [摄氏度] / the float zero sentinel *)
    DL_SIP_TTIMEZERO : TIME := T#0S;        (* 零时长哨兵 [ms] / the zero duration sentinel *)
    DL_SIP_MS_SEC    : DINT := 1000;        (* 毫秒到秒常量除子（R382 级联口径）[ms/s] / the constant milliseconds per second divisor *)
    DL_SIP_ZERO      : UDINT := 0;          (* 无符号零哨兵 [码或秒或次] / the unsigned zero sentinel *)
    DL_SIP_ONE       : UDINT := 1;          (* 计数步进 [次] / the count step *)
    DL_SIP_CMAX      : UDINT := 2147483000; (* 扰动计数饱和上限（防回绕）[次] / the disturbance count saturation cap *)
END_VAR

// 段 0｜复位沿无条件调用（规则 ⑦）/ segment 0, the unconditional reset edge refresh
rtReset(CLK := bReset);                    // 每拍无条件刷新 / refreshed every scan

// 段 1｜首拍初始化与出口内部位预清（R310 / R256）/ segment 1, the first scan init and the presets
IF NOT _bInit THEN                         // 首拍一拍 / the first scan
    _bInit := TRUE;                        // 置首拍标志 / raise the first scan flag
    _bFault := FALSE;                      // 故障锁存显式清零 / clear the fault latch explicitly
    _eState := E_DL_SipPhase.eIdle;        // 状态显式落空闲 / place the state to idle
END_IF

// 段 2｜域闸（R272 全枚举：fTempC 非有限闸 + fHoldTempSet 非有限与承诺段闸）/ segment 2, the domain gates
_bTInBad := (fTempC <> fTempC) OR ((fTempC - fTempC) <> DL_SIP_TZERO); // 温度非有限（R79 双判）/ the temperature non finite
_bCfgBad := (fHoldTempSet <> fHoldTempSet) OR ((fHoldTempSet - fHoldTempSet) <> DL_SIP_TZERO) // 设定非有限 / the setpoint non finite
         OR (fHoldTempSet < DL_SIP_TSETMIN) // 设定越承诺段下界 / the setpoint under the promise
         OR (tHoldTime <= DL_SIP_TTIMEZERO) // 保温窗非正 / a non positive hold window
         OR (tDrainTimeout <= DL_SIP_TTIMEZERO); // 排凝超时非正 / a non positive drain timeout

// 段 3｜本拍实时温度判据（R42：迁入与驻留判温均取本拍值；NaN 不许当冷值漏判）/ segment 3, the live temperature verdict
IF (NOT _bTInBad) AND (NOT _bCfgBad) THEN  // 双闸通过才判 / both gates passed
    _bTempOk := fTempC >= fHoldTempSet;    // 达标本拍实时值 / the live verdict
ELSE                                       // 闸未通过 / the gates failed
    _bTempOk := FALSE;                     // 达标判据强制假（安全侧）/ force the verdict false
END_IF

// 段 4｜复位沿与首次成因锁存（复位沿唯一解除，R188；故障期不重推断，R189；组态根因优先）/ segment 4, the reset edge and the first cause latch
IF rtReset.Q THEN                          // 复位上升沿 / the reset rising edge
    _bFault := FALSE;                      // 清故障锁存（恒可达，R152 自证）/ clear the fault latch
    _nCodeLatch := DL_SIP_ZERO;            // 清锁存码 / clear the latched code
    _eState := E_DL_SipPhase.eIdle;        // 迁回空闲 / back to idle
    _bReleased := FALSE;                   // 清放行内部锁存（批界复位）/ clear the release latch
    uDisturbCount := DL_SIP_ZERO;          // 清扰动计数（批次台账随批清，作用域声明边界九）/ clear the disturbance count
END_IF
IF NOT _bFault THEN                        // 未锁存才登记成因 / register only while not latched
    IF _bCfgBad THEN                       // 组态非法（根因优先归因）/ the config fault first
        _bFault := TRUE;                   // 置锁存 / latch
        _nCodeLatch := DL_SIP_CODE_SET;    // 登记设定码 / register the setpoint code
        IF (tHoldTime <= DL_SIP_TTIMEZERO) OR (tDrainTimeout <= DL_SIP_TTIMEZERO) THEN // 时间组态单独归因（R190 成因独立码）/ the time config attribution
            _nCodeLatch := DL_SIP_CODE_TIME; // 登记时间码 / register the time code
        END_IF
    ELSIF _bTInBad THEN                    // 温度非有限（状态不明不得放行，直接锁存）/ the probe fault
        _bFault := TRUE;                   // 置锁存 / latch
        _nCodeLatch := DL_SIP_CODE_TEMP;   // 登记探头码 / register the probe code
    END_IF
END_IF

// 段 5｜主状态机（ENUM + CASE，ELSE 兜底；迁入安全相带全量闸位复检，R274）/ segment 5, the main state machine
CASE _eState OF

    E_DL_SipPhase.eIdle:                   // 空闲相 / the idle phase
        _bDrain := FALSE;                  // 双输出内部位清零（R57）/ clear the internal bits
        _bSteam := FALSE;                  // 双输出内部位清零 / clear the internal bits
        IF bEn AND (NOT _bFault) AND (NOT _bCfgBad) THEN // 使能 ∧ 组态闸（迁入闸位复检，R274）/ the start gate
            _eState := E_DL_SipPhase.eDrain; // 迁入排凝相 / enter the drain phase
        END_IF

    E_DL_SipPhase.eDrain:                  // 排凝相：开排凝等反馈 / the drain phase
        _bDrain := TRUE;                   // 排凝指令 / the drain command
        _bSteam := FALSE;                  // 蒸汽关断 / the steam off
        // 失能或温度失效不在此自行迁出：由段 4 首次成因锁存 + 段 5b 统一迁入闸接管。
        // A disable or a probe loss does not exit here, the unified gates take over.
        IF bDrainDone THEN                 // 排凝完成反馈 / the drain done feedback
            _bDrain := FALSE;              // 撤排凝 / drop the drain command
            _eState := E_DL_SipPhase.eHeatUp; // 迁入升温相 / enter the heat up phase
        ELSIF tonDrain.Q THEN              // 排凝超时（看门狗到时）/ the drain timeout
            _bFault := TRUE;               // 置锁存 / latch the fault
            _nCodeLatch := DL_SIP_CODE_DRAIN; // 登记超时码 / register the timeout code
        END_IF

    E_DL_SipPhase.eHeatUp:                 // 升温相：开蒸汽等达标（本拍实时判温，R42）/ the heat up phase
        _bDrain := FALSE;                  // 排凝撤 / drop the drain
        _bSteam := TRUE;                   // 蒸汽开 / the steam on
        IF _bTInBad THEN                   // 温度失效（关断由故障路径统一执行）/ the probe loss
            _bFault := TRUE;               // 置锁存 / latch
            _nCodeLatch := DL_SIP_CODE_TEMP; // 登记探头码 / register the probe code
        ELSIF _bTempOk THEN                // 本拍达标（实时值，无跨拍陈旧判据）/ the live verdict
            _eState := E_DL_SipPhase.eHold; // 迁入保温相（迁入拍即计时使能）/ enter the hold phase
        END_IF

    E_DL_SipPhase.eHold:                   // 保温相：TON 计时，跌破重计（断点重计口径）/ the hold phase
        _bSteam := TRUE;                   // 蒸汽保持 / the steam holds
        IF _bTInBad THEN                   // 温度失效 / the probe loss
            _bFault := TRUE;               // 置锁存 / latch
            _nCodeLatch := DL_SIP_CODE_TEMP; // 登记探头码 / register the probe code
        ELSIF NOT _bTempOk THEN            // 跌破设定（本拍实时值）：计时中止回升温 + 扰动计数 / the drop below setpoint
            IF uDisturbCount < DL_SIP_CMAX THEN // 饱和闸（防回绕）/ the saturation cap
                uDisturbCount := uDisturbCount + DL_SIP_ONE; // 扰动计数 + 1 / count the disturbance
            END_IF
            _eState := E_DL_SipPhase.eHeatUp; // 回升温相（TON IN 随相撤自动清零重计）/ back to heat up
        ELSIF tonHold.Q THEN               // 保温窗计满（连续无跌破）/ the window elapsed
            _bSteam := FALSE;              // 关蒸汽 / the steam off
            _eState := E_DL_SipPhase.eCooldown; // 迁入冷却相 / enter the cooldown phase
        END_IF

    E_DL_SipPhase.eCooldown:               // 冷却相：关蒸汽等回落确认 / the cooldown phase
        _bSteam := FALSE;                  // 蒸汽关断 / the steam off
        IF _bTInBad THEN                   // 温度失效 / the probe loss
            _bFault := TRUE;               // 置锁存 / latch
            _nCodeLatch := DL_SIP_CODE_TEMP; // 登记探头码 / register the probe code
        ELSIF NOT _bTempOk THEN            // 回落确认（复用本拍达标判据的补集，双闸已过才可比）/ the fall below confirmed
            _bReleased := TRUE;            // 放行内部锁存 / latch the release
            _eState := E_DL_SipPhase.eDone; // 迁入完成相 / enter the done phase
        END_IF

    E_DL_SipPhase.eDone:                   // 完成相：bSterilized 保持（批界清除）/ the done phase
        _bSteam := FALSE;                  // 蒸汽保持关断 / the steam off
        IF NOT bEn THEN                    // 批界：失能（复位沿已由段 4 先行处理）/ the batch boundary on disable
            _bReleased := FALSE;           // 清放行 / clear the release
            _eState := E_DL_SipPhase.eIdle; // 迁回空闲 / back to idle
        END_IF

    E_DL_SipPhase.eFault:                  // 故障相：双输出关断等复位沿 / the fault phase
        _bDrain := FALSE;                  // 排凝关断 / the drain off
        _bSteam := FALSE;                  // 蒸汽关断（安全侧）/ the steam off
        _bReleased := FALSE;               // 放行撤销（故障期不放行）/ the release withdrawn
        IF NOT _bFault THEN                // 锁存已清才迁出 / the exit after the latch cleared
            _eState := E_DL_SipPhase.eIdle; // 迁回空闲 / back to idle
        END_IF

    ELSE                                   // 非法枚举值拦截 / the illegal enumeration guard
        _eState := E_DL_SipPhase.eFault;   // 落故障相 / force to the fault phase
        _bFault := TRUE;                   // 置锁存 / latch the fault
        _nCodeLatch := DL_SIP_CODE_TEMP;   // 复用温度码（R90 反证：非法枚举不可达无独立观测需求）/ reuse the probe code

END_CASE

// 段 5b｜故障统一迁入闸（置于状态机之后，R274 迁入完备性）/ segment 5b, the unified fault entry gate
IF _bFault AND (_eState <> E_DL_SipPhase.eFault) THEN // 已锁存但不在故障相 / latched but not in the fault phase
    _eState := E_DL_SipPhase.eFault;       // 任何相检出故障一律落故障相 / any phase with a latch lands in the fault phase
END_IF

// 段 5c｜失能停机相输出清零（锁存保留，R57 / R191 声明；eDone 批界已自处理）/ segment 5c, the disable clearing
IF (NOT bEn) AND (_eState <> E_DL_SipPhase.eFault) AND (_eState <> E_DL_SipPhase.eDone) THEN // 失能且不在故障 / 完成相 / disabled
    _eState := E_DL_SipPhase.eIdle;        // 撤工艺回空闲 / back to idle
    _bDrain := FALSE;                      // 双输出清零 / clear the bits
    _bSteam := FALSE;                      // 双输出清零 / clear the bits
    _bReleased := FALSE;                   // 放行撤销 / the release withdrawn
END_IF

// 段 6｜双定时器无条件调用（IN 为相驻留显式条件；tonHold IN 含本拍达标判据，跌破即断计重计）/ segment 6, the unconditional timers
tonDrain(IN := (_eState = E_DL_SipPhase.eDrain) AND bEn AND (NOT _bFault), PT := tDrainTimeout); // 排凝看门狗 / the drain watchdog
tonHold(IN := (_eState = E_DL_SipPhase.eHold) AND _bTempOk AND bEn AND (NOT _bFault), PT := tHoldTime); // 保温计时（跌破即断计）/ the hold timer

// 段 7｜保温剩余倒计时（非保温相为 0；常量除子 1000，零除法面）/ segment 7, the hold remaining countdown
IF _eState = E_DL_SipPhase.eHold THEN      // 保温相内计算 / inside the hold phase
    nRemainMs := TIME_TO_DINT(tHoldTime) - TIME_TO_DINT(tonHold.ET); // 剩余毫秒 / the remaining milliseconds
    IF nRemainMs < 0 THEN                  // 负值防御（饱和为零）/ the negative guard
        nRemainMs := 0;                    // 钳到零 / clamp to zero
    END_IF
    uHoldRemain := DINT_TO_UDINT(nRemainMs / DL_SIP_MS_SEC); // 常量除子秒化 / the constant divisor seconds
ELSE                                       // 非保温相 / the other phases
    uHoldRemain := DL_SIP_ZERO;            // 倒计时清零 / zero the countdown
END_IF

// 段 8｜统一出口（名实双出口同源，R191）/ segment 8, the unified outlet
bDrainCmd := _bDrain AND bEn AND (NOT _bFault); // 排凝出口（失能 / 故障双保险）/ the drain outlet
bSteamCmd := _bSteam AND bEn AND (NOT _bFault); // 蒸汽出口（安全侧关断双保险）/ the steam outlet
bSterilized := _bReleased AND (NOT _bFault); // 放行出口（故障期撤销）/ the release outlet
eState := _eState;                         // 状态出口 / the state outlet
bError := _bFault;                         // 故障标志与锁存同源 / the fault flag from the latch
IF _bFault THEN                            // 故障锁存回放（R187）/ the latched replay
    nErrCode := _nCodeLatch;               // 回放锁存码 / replay the latched code
ELSE                                       // 无事件 / no event
    nErrCode := DL_SIP_ZERO;               // 正常 / ok
END_IF
END_FUNCTION_BLOCK

(* ---- FB_DL_SolarStringGroundFault.st ---- *)
//==============================================================================
// 功能块：FB_DL_SolarStringGroundFault ｜ 中文名称：光伏组串对地绝缘阻抗检测
// 所属子库：DL_Process ｜ 版本：v1.0.1 ｜ 兼容：CODESYS V3.5+ / TwinCAT 3 / 汇川 InoProShop
// 功能描述：光伏组串对地绝缘阻抗检测（不平衡电桥法）：由正/负母线对地电压与组串母线
//           电压推算正极、负极与并联对地绝缘电阻，按两级阈值告警（确认拍数 + 锁存）。
//           本件仅监视不控：不触发脱扣、不切组串、不做绝缘老化趋势记录（趋势归上位）。
// 开源溯源 (Origin)：道莅原创实现（参考 不平衡电桥法公开测量原理 分类与参数域）
// 单位表：母线及对地电压[V] / 绝缘电阻与桥阻[kΩ] / 阈值[kΩ] / 确认拍数[拍] /
//         失衡比值[无量纲] / 电压判零容差[V]
// ------------------------------------------------------------------------------
// 量纲链（R108 量纲组合表，编码前逐式复核，禁凭记忆落码）：
//   设 Gp = 1/Rp、Gn = 1/Rn 分别为正/负母线对地漏电导，G_t = Gp + Gn 为总漏电导，
//   Rb 为测量桥阻。桥阻上的压降为 (Vbus − Vp − Vn)，其上电流即总漏电流：
//     G_t [1/kΩ] = (Vbus − Vp − Vn) / (Rb × (Vp + Vn))        —— 量纲：V/(kΩ·V) = 1/kΩ
//   两端漏电按对地电压分压比分配（同一漏电网络的基尔霍夫关系）：
//     Gp / Gn = Vn / Vp   →   Gp = G_t × Vn/(Vp+Vn)，Gn = G_t × Vp/(Vp+Vn)
//   取倒数得电阻（kΩ）：
//     R_t = 1/G_t = Rb × (Vp + Vn) / (Vbus − Vp − Vn)
//     Rp  = R_t × (Vp + Vn) / Vn
//     Rn  = R_t × (Vp + Vn) / Vp
//   复核：Rp/Rn = Vp/Vn（与电桥分压比一致）；并联合成 1/(1/Rp + 1/Rn) = R_t（自洽）。
//   注意（本件最高风险点）：R_t 的除子为 (Vbus − Vp − Vn)。当组串绝缘趋于无穷（正负
//   完全平衡、Vp + Vn 逼近 Vbus）时 R_t 趋于无穷；此时若照抄「Rb × (Vbus/(Vp+Vn) − 1)」
//   这种乘式写法，会得到趋于 0 的伪阻值（量纲虽为 kΩ，物理上却是倒数关系），从而把
//   绝缘良好误判成对地短路并误告警。本件一律用除式，并对「完全平衡退化」给出显式分支：
//   (Vbus − Vp − Vn) ≤ 1.0 V 时判为绝缘无穷大，取上限哨兵 1.0E9 kΩ 输出、不告警、
//   不计告警确认拍数（不冒充实测值，HMI 以饱和值显示）。
// ------------------------------------------------------------------------------
// 错误码表：16#0005_0410 信息级（母线电压 ≤ 0，或 Vp + Vn 近零，或单极对地电压非正：
//           绝缘推算不可判，禁止输出伪阻值，bUndecidable 置位，不置 bError）/
//           16#0005_0411 信息级（单极对地阻抗失衡提示：max(Rp,Rn)/min(Rp,Rn) > 3，
//           不置 bError）/ 16#0005_035A 故障级（桥阻非正或告警阈值倒置，置 bError）/
//           16#0005_035B 故障级（输入非有限，置 bError，阻值输出回零）/ 16#0005_035C
//           故障级兜底（状态机落 ELSE 非法状态，置 bError）。码位 16#0005 段。
// 状态机：E_DL_StringInsState（eIdle=0 待机 / eMeasure=10 正常推算 / eUndecidable=20
//           推算不可判 / eAlarm=30 告警锁存后监视 / eFault=99 故障兜底），CASE 含 ELSE
//           兜底，ELSE 置 035C 且阻值回零、许可撤。
// 边界行为：① 量纲链见上（除式 + 完全平衡退化显式分支）；② Vp + Vn ≤ 1.0 V 或
//           fBusV ≤ 0 → 信息 0410 + bUndecidable := TRUE + bValid := FALSE（推算不可判
//           时禁止输出伪阻值）；单极对地电压非正同理（分压比不可算）；③ fBridgeKOhm ≤ 0
//           或 fAlarmKOhm ≥ fWarnKOhm → 故障 035A；④ 非有限（NaN 自反判 + Inf 幅值上限
//           判）→ 故障 035B，阻值回零；⑤ 分级：R_t < 告警阈值 → bAlarm；R_t < 预警阈值
//           → bWarn；均需连续 nConfirmSamples 拍确认，确认后锁存至 bReset（防单点误报
//           停机）；⑥ 失衡判据 max/min > 3.0（常量），命中即 bUnbalanced + 信息 0411；
//           ⑦ 失能 → 不判、bValid := FALSE，但绝不清除已锁存的 bWarn/bAlarm（告警是
//           历史事实，只能人工复位）。
// 验收向量（算法已证，手算）：① Vbus = 600 V、Vp = 300 V、Vn = 300 V、Rb = 100 kΩ →
//           Vbus − Vp − Vn = 0 → 完全平衡退化分支 → R_t = 1.0E9 kΩ 哨兵、bWarn/bAlarm
//           均为 FALSE（若用乘式写法此处会得 0 kΩ 并误告警，本向量即该风险的回归用例）；
//           ② Vbus = 600 V、Vp = 310 V、Vn = 290 V、Rb = 100 kΩ → Vbus − Vp − Vn = 0 V
//           仍属退化（差值阈值内）→ 同样取 1.0E9 kΩ 上限哨兵；改取 Vp = 310 V、Vn = 280 V（差 10 V）→
//           R_t = 100 × 590 / 10 = 5900 kΩ、Rp = 5900 × 590/280 ≈ 12432 kΩ、
//           Rn = 5900 × 590/310 ≈ 11229 kΩ，失衡比 1.11 < 3 → 不告警不失衡；
//           ③ 阈值 告警 100、预警 1000 kΩ，实测 R_t = 80 kΩ → 连续 3 拍确认 → bAlarm
//           锁存；④ Vp + Vn = 0.5 V → 信息 0410 + bUndecidable + bValid := FALSE。
//           编译器已证（三平台）：未跑，由收口方登记。
// 修订历史：v1.0.0 2026-11-17 首版（R25 派单 · §4.20）
//           v1.0.1 2026-11-17 终审补域端点闸（对外引脚契约零变更）：预警阈值 fWarnKOhm 若被配到
//           ≥ 上限哨兵 DL_SGF_R_MAX（1.0E9 kΩ），完全平衡退化分支输出的哨兵值会被判为「低于预警阈值」
//           而误报警（把绝缘良好判成异常）。组态闸补一项 fWarnKOhm >= DL_SGF_R_MAX → 035A。
//           总监独立验算裁定：派单书 §4.20 的乘式 Rb x (Vbus/(Vp+Vn) − 1) 分子分母倒置（完全平衡
//           时得 0 kΩ、单极短路时得无穷），本件除式 Rb x (Vp+Vn)/(Vbus − Vp − Vn) 在两端均取正确
//           极限（D→0 ⇒ R→∞；Vp+Vn→0 ⇒ R→0），编码侧改法正确，派单书须勘误。
//==============================================================================
(*------------------------------------------------------------------------------
 * 枚举: E_DL_StringInsState（归属 DL_Process，与 FB_DL_SolarStringGroundFault 同文件）
 *----------------------------------------------------------------------------*)
TYPE E_DL_StringInsState :
(
    eIdle        := 0,   // 待机：失能，不推算不判定 / Idle, neither computed nor judged
    eMeasure     := 10,  // 正常推算：阻值有效 / Normal measurement, valid resistances
    eUndecidable := 20,  // 推算不可判：母线或对地电压条件不成立 / Undecidable, the voltage conditions do not hold
    eAlarm       := 30,  // 告警锁存后监视：阻值仍有效 / Monitoring after a latched alarm
    eFault       := 99   // 故障兜底：组态非法/非有限/非法状态 / Fault fallback
);
END_TYPE

(*==============================================================================
 * 功能块: FB_DL_SolarStringGroundFault
 * 调用约定: 每个扫描周期无条件调用一次；电压量由直流侧采样与滤波层刷新。
 *============================================================================*)
FUNCTION_BLOCK FB_DL_SolarStringGroundFault
VAR_INPUT
    fPosToGroundV   : LREAL;                       // 正母线对地电压 [V] / Positive bus voltage to ground [V]
    fNegToGroundV   : LREAL;                       // 负母线对地电压（幅值）[V] / Negative bus voltage to ground, magnitude [V]
    fBusV           : LREAL;                       // 组串母线电压 [V]，须 > 0 / String bus voltage [V], must be > 0
    fBridgeKOhm     : LREAL := 100.0;              // 测量桥电阻 [kΩ]，须 > 0 / Measurement bridge resistance [kΩ], must be > 0
    fWarnKOhm       : LREAL := 1000.0;             // 预警阈值 [kΩ] / Warning threshold [kΩ]
    fAlarmKOhm      : LREAL := 100.0;              // 告警阈值 [kΩ]，须 < 预警阈值 / Alarm threshold [kΩ], must be below the warning
    nConfirmSamples : INT := 3;                    // 告警确认拍数 [拍]，域 1~20 / Alarm confirmation samples, domain 1..20
    bEnable         : BOOL;                        // 总使能 / Master enable
    bReset          : BOOL;                        // 复位，上升沿清告警锁存 / Reset, rising edge clears the latched alarms
END_VAR
VAR_OUTPUT
    fInsPosKOhm     : LREAL;                       // 正极对地绝缘电阻 [kΩ] / Positive-to-ground insulation resistance [kΩ]
    fInsNegKOhm     : LREAL;                       // 负极对地绝缘电阻 [kΩ] / Negative-to-ground insulation resistance [kΩ]
    fInsTotalKOhm   : LREAL;                       // 并联对地绝缘电阻 [kΩ] / Parallel insulation resistance [kΩ]
    bWarn           : BOOL;                        // 预警（确认后锁存至 bReset）/ Warning, latched until reset after confirmation
    bAlarm          : BOOL;                        // 告警（确认后锁存至 bReset）/ Alarm, latched until reset after confirmation
    bUnbalanced     : BOOL;                        // 正负极失衡（max/min > 3）/ Positive-negative imbalance
    bUndecidable    : BOOL;                        // 推算不可判（禁止使用阻值输出）/ Undecidable, the resistance outputs must not be used
    eErr            : UDINT;                       // 错误码，0 = 无错，码位 16#0005_0410 起信息级、16#0005_035A 起故障级（分带见错误码表） / Error code, 0 = no error, band info/fault per the code table
    bError          : BOOL;                        // 故障级标志，仅故障级错误置位 / Fault-class flag, set only on fault-level codes
    bValid          : BOOL;                        // 阻值输出可用标志，不可判/失能/故障闸显式 FALSE / Resistance usable flag, explicit FALSE when undecidable, disabled or faulted
    eState          : E_DL_StringInsState;         // 主状态机当前状态 / Current state of the main state machine
END_VAR
VAR
    fbReset         : R_TRIG;                      // 复位上升沿检测实例 / Reset rising edge detector
    fSumV           : LREAL;                       // 对地电压之和 Vp + Vn [V] / Sum of the ground voltages [V]
    fDiffV          : LREAL;                       // 母线电压盈余 Vbus − (Vp + Vn) [V] / Bus voltage surplus [V]
    fTotalKOhm      : LREAL;                       // 并联绝缘电阻工作值 [kΩ] / Parallel insulation working value [kΩ]
    fPosKOhm        : LREAL;                       // 正极绝缘电阻工作值 [kΩ] / Positive insulation working value [kΩ]
    fNegKOhm        : LREAL;                       // 负极绝缘电阻工作值 [kΩ] / Negative insulation working value [kΩ]
    fRatio          : LREAL;                       // 失衡比值 max/min [无量纲] / Imbalance ratio max/min
    fMaxKOhm        : LREAL;                       // 两极大值 [kΩ] / Maximum of both poles [kΩ]
    fMinKOhm        : LREAL;                       // 两极小值 [kΩ] / Minimum of both poles [kΩ]
    nConfirmEff     : INT;                         // 钳位后的确认拍数 [拍] / Clamped confirmation samples
    nWarnCnt        : INT;                         // 预警连续确认计数 [拍] / Consecutive warning samples
    nAlarmCnt       : INT;                         // 告警连续确认计数 [拍] / Consecutive alarm samples
    bNonFin         : BOOL;                        // 非有限判定中间标志 / Non-finite detection intermediate flag
    bUndecidableNow : BOOL;                        // 本拍不可判标志 / Undecidable this scan
    bDegenerate     : BOOL;                        // 完全平衡退化标志 / Fully balanced degenerate case
    bWarnNow        : BOOL;                        // 本拍预警判据 / Warning predicate this scan
    bAlarmNow       : BOOL;                        // 本拍告警判据 / Alarm predicate this scan
    bFirstScan      : BOOL := TRUE;                // 上电首拍标志 / First-scan flag
END_VAR
VAR CONSTANT
    DL_SGF_CODE_INFO_1 : UDINT := 16#0005_0410;    // 信息级槽 1（推算不可判） / info slot 1
    DL_SGF_CODE_INFO_2 : UDINT := 16#0005_0411;    // 信息级槽 2（单极对地阻抗失衡提示） / info slot 2
    DL_SGF_CODE_FLT_1  : UDINT := 16#0005_035A;    // 故障级槽 1（桥阻/阈值组态非法） / fault slot 1
    DL_SGF_CODE_FLT_2  : UDINT := 16#0005_035B;    // 故障级槽 2（输入非有限） / fault slot 2
    DL_SGF_CODE_FLT_3  : UDINT := 16#0005_035C;    // 故障级槽 3（非法状态兜底） / fault slot 3
    DL_SGF_R_MAX       : LREAL := 1.0E9;           // 绝缘电阻上限哨兵（完全平衡退化取值）[kΩ] / Insulation ceiling sentinel [kΩ]
    DL_SGF_VMIN        : LREAL := 1.0;             // 对地电压和与母线盈余判零门限 [V] / Voltage sum and surplus threshold [V]
    DL_SGF_IMB_RATIO   : LREAL := 3.0;             // 失衡比值门限 [无量纲] / Imbalance ratio threshold
    DL_SGF_CONF_MIN    : INT := 1;                 // 确认拍数下限 [拍] / Confirmation floor [samples]
    DL_SGF_CONF_MAX    : INT := 20;                // 确认拍数上限 [拍] / Confirmation ceiling [samples]
    DL_SGF_ZERO        : LREAL := 0.0;             // 零值常量，避免裸字面量 [—] / Zero constant, avoids a bare literal
    DL_SGF_TOL         : LREAL := 1.0E-6;          // 浮点比较容差 [—] / Float comparison tolerance
    DL_SGF_INF         : LREAL := 1.7976931348623157E308; // LREAL 幅值上限，Inf 判据 / LREAL magnitude ceiling
END_VAR

(*------------------------------------------------------------------------------
 * 段 1｜无条件刷新区（红线 5）：复位沿检测在任意分支之外周期调用
 *----------------------------------------------------------------------------*)
fbReset(CLK := bReset);                            // 复位沿检测无条件刷新 / reset edge refreshed unconditionally

(*------------------------------------------------------------------------------
 * 段 2｜复位沿处理（改写置于沿后，防吞沿 R39）：清告警锁存与确认计数
 *----------------------------------------------------------------------------*)
IF fbReset.Q THEN
    eState := E_DL_StringInsState.eIdle;
    eErr   := 16#0000_0000;                        // 复位清码 / reset clears the code
    bError := FALSE;                               // 复位清故障 / reset clears the fault
    bWarn  := FALSE;                               // 预警锁存清（仅人工复位可清）/ warning latch cleared
    bAlarm := FALSE;                               // 告警锁存清（仅人工复位可清）/ alarm latch cleared
    nWarnCnt := 0;                                 // 预警确认计数清 / warning counter cleared
    nAlarmCnt := 0;                                // 告警确认计数清 / alarm counter cleared
    bFirstScan := TRUE;                            // 重新首拍化 / re-initialize first scan
END_IF

(*------------------------------------------------------------------------------
 * 段 3｜非有限输入闸：035B + 阻值回零（故障路径输出安全值而非上次值，红线 6）
 *----------------------------------------------------------------------------*)
bNonFin := (fPosToGroundV <> fPosToGroundV) OR (ABS(fPosToGroundV) >= DL_SGF_INF)
        OR (fNegToGroundV <> fNegToGroundV) OR (ABS(fNegToGroundV) >= DL_SGF_INF)
        OR (fBusV <> fBusV) OR (ABS(fBusV) >= DL_SGF_INF)
        OR (fBridgeKOhm <> fBridgeKOhm) OR (ABS(fBridgeKOhm) >= DL_SGF_INF)
        OR (fWarnKOhm <> fWarnKOhm) OR (ABS(fWarnKOhm) >= DL_SGF_INF)
        OR (fAlarmKOhm <> fAlarmKOhm) OR (ABS(fAlarmKOhm) >= DL_SGF_INF);   // 引脚非有限汇总 / pins non-finite
IF bNonFin THEN
    eState := E_DL_StringInsState.eFault;          // 进故障相 / enter fault state
    eErr   := DL_SGF_CODE_FLT_2;                   // 故障级：输入非有限 / fault: non-finite input
    bError := TRUE;                                // 故障级必置 bError（R45 配对）/ fault-class pairs with bError
    bValid := FALSE;                               // 阻值不可用 / resistances unusable
    fInsPosKOhm := DL_SGF_ZERO;                    // 正极阻值回零安全侧 / positive resistance zeroed, safe side
    fInsNegKOhm := DL_SGF_ZERO;                    // 负极阻值回零安全侧 / negative resistance zeroed, safe side
    fInsTotalKOhm := DL_SGF_ZERO;                  // 并联阻值回零安全侧 / parallel resistance zeroed, safe side
    bUnbalanced := FALSE;                          // 失衡标志撤 / imbalance withdrawn
    bUndecidable := FALSE;                         // 不可判标志撤（故障优先）/ undecidable withdrawn, fault outranks
    RETURN;
END_IF

(*------------------------------------------------------------------------------
 * 段 4｜组态合法性闸：桥阻须为正（否则除零）、告警阈值须严格小于预警阈值
 *----------------------------------------------------------------------------*)
IF (fBridgeKOhm <= DL_SGF_TOL) OR (fAlarmKOhm >= fWarnKOhm - DL_SGF_TOL)
   OR (fWarnKOhm >= DL_SGF_R_MAX) THEN
    eState := E_DL_StringInsState.eFault;          // 进故障相 / enter fault state
    eErr   := DL_SGF_CODE_FLT_1;                   // 故障级：桥阻/阈值组态非法 / fault: bridge or threshold configuration invalid
    bError := TRUE;                                // 故障级必置 bError（R45 配对）/ fault-class pairs with bError
    bValid := FALSE;                               // 阻值不可用 / resistances unusable
    fInsPosKOhm := DL_SGF_ZERO;                    // 正极阻值回零安全侧 / positive resistance zeroed
    fInsNegKOhm := DL_SGF_ZERO;                    // 负极阻值回零安全侧 / negative resistance zeroed
    fInsTotalKOhm := DL_SGF_ZERO;                  // 并联阻值回零安全侧 / parallel resistance zeroed
    bUnbalanced := FALSE;                          // 失衡标志撤 / imbalance withdrawn
    bUndecidable := FALSE;                         // 不可判标志撤 / undecidable withdrawn
    RETURN;
END_IF

(*------------------------------------------------------------------------------
 * 段 5｜组态钳位：确认拍数钳到 1~20（域外按边界钳，不新占码位）
 *----------------------------------------------------------------------------*)
nConfirmEff := nConfirmSamples;                    // 先取引脚值 / take the pin value first
IF nConfirmEff < DL_SGF_CONF_MIN THEN
    nConfirmEff := DL_SGF_CONF_MIN;                // 下限钳位 [拍] / clipped to the floor
END_IF
IF nConfirmEff > DL_SGF_CONF_MAX THEN
    nConfirmEff := DL_SGF_CONF_MAX;                // 上限钳位 [拍] / clipped to the ceiling
END_IF

(*------------------------------------------------------------------------------
 * 段 6｜不可判闸（R42 家族：推算不成立时禁止输出伪阻值）：
 *       母线电压 ≤ 0、对地电压和近零、或任一极对地电压非正 → 0410 + bUndecidable
 *       此时阻值输出回零且 bValid := FALSE，绝不给出"看起来能信"的数字
 *----------------------------------------------------------------------------*)
fSumV := fPosToGroundV + fNegToGroundV;            // 对地电压之和 [V] / sum of the ground voltages [V]
bUndecidableNow := (fBusV <= DL_SGF_TOL)
                OR (fSumV <= DL_SGF_VMIN)
                OR (fPosToGroundV <= DL_SGF_TOL)
                OR (fNegToGroundV <= DL_SGF_TOL);  // 不可判判据（四项任一）/ undecidable predicate
IF bUndecidableNow THEN
    bUndecidable := TRUE;                          // 不可判标志置位 / undecidable raised
    bValid := FALSE;                               // 阻值不可用（禁伪阻值）/ resistances unusable
    fInsPosKOhm := DL_SGF_ZERO;                    // 正极阻值回零 / positive resistance zeroed
    fInsNegKOhm := DL_SGF_ZERO;                    // 负极阻值回零 / negative resistance zeroed
    fInsTotalKOhm := DL_SGF_ZERO;                  // 并联阻值回零 / parallel resistance zeroed
    bUnbalanced := FALSE;                          // 不可判时不判失衡 / no imbalance verdict when undecidable
    nWarnCnt := 0;                                 // 确认计数清零（不可判拍不计入）/ confirmation counters cleared
    nAlarmCnt := 0;
    bWarnNow := FALSE;                             // 本拍不出判据 / no predicate this scan
    bAlarmNow := FALSE;
    eState := E_DL_StringInsState.eUndecidable;    // 进不可判相 / enter the undecidable state
    eErr := DL_SGF_CODE_INFO_1;                    // 信息级：绝缘推算不可判 / info: insulation not decidable
    bError := FALSE;                               // 信息级不置 bError（R45/R101）/ info never raises bError
ELSE
    (*--------------------------------------------------------------------------
     * 段 7｜量纲链落码（除式，禁乘式）：R_t = Rb x (Vp + Vn) / (Vbus − Vp − Vn)
     *   完全平衡退化（Vbus − Vp − Vn ≤ 1.0 V，绝缘趋无穷）→ 显式取上限哨兵，
     *   绝不让除子趋零、也绝不用乘式（乘式会把无穷绝缘算成 0 kΩ 并误告警）
     *-------------------------------------------------------------------------*)
    bDegenerate := FALSE;                          // 退化标志初值 / degenerate seed
    fDiffV := fBusV - fSumV;                       // 母线盈余 [V] / bus surplus [V]
    IF fDiffV <= DL_SGF_VMIN THEN
        bDegenerate := TRUE;                       // 完全平衡退化分支（显式）/ explicit degenerate branch
        fTotalKOhm := DL_SGF_R_MAX;                // 绝缘取上限哨兵 [kΩ] / insulation takes the ceiling sentinel
        fPosKOhm := DL_SGF_R_MAX;                  // 正极阻值同为上限哨兵 [kΩ] / positive takes the ceiling sentinel
        fNegKOhm := DL_SGF_R_MAX;                  // 负极阻值同为上限哨兵 [kΩ] / negative takes the ceiling sentinel
    ELSE
        fTotalKOhm := fBridgeKOhm * fSumV / fDiffV;                      // 并联绝缘电阻 [kΩ] / parallel insulation [kΩ]
        IF fTotalKOhm > DL_SGF_R_MAX THEN
            fTotalKOhm := DL_SGF_R_MAX;            // 上限饱和（防溢出）[kΩ] / ceiling saturation
        END_IF
        fPosKOhm := fTotalKOhm * fSumV / fNegToGroundV;                  // 正极 = R_t x (Vp+Vn)/Vn（除子段 6 已判非零）[kΩ] / positive pole
        fNegKOhm := fTotalKOhm * fSumV / fPosToGroundV;                  // 负极 = R_t x (Vp+Vn)/Vp [kΩ] / negative pole
        IF fPosKOhm > DL_SGF_R_MAX THEN
            fPosKOhm := DL_SGF_R_MAX;              // 上限饱和 [kΩ] / ceiling saturation
        END_IF
        IF fNegKOhm > DL_SGF_R_MAX THEN
            fNegKOhm := DL_SGF_R_MAX;              // 上限饱和 [kΩ] / ceiling saturation
        END_IF
    END_IF
    fInsPosKOhm := fPosKOhm;                       // 正极阻值出口 [kΩ] / positive resistance outlet
    fInsNegKOhm := fNegKOhm;                       // 负极阻值出口 [kΩ] / negative resistance outlet
    fInsTotalKOhm := fTotalKOhm;                   // 并联阻值出口 [kΩ] / parallel resistance outlet
    bUndecidable := FALSE;                         // 推算成立：不可判标志撤 / decidable, the flag drops
    bValid := TRUE;                                // 阻值可用 / resistances usable
    bError := FALSE;                               // 推算路径无故障 / no fault on the measurement path

    (*--------------------------------------------------------------------------
     * 段 8｜失衡判据：max(Rp,Rn) / min(Rp,Rn) > 3.0（除子先判零，退化时比值记 1）
     *-------------------------------------------------------------------------*)
    fMaxKOhm := fPosKOhm;                          // 极大值种子 / maximum seed
    IF fNegKOhm > fMaxKOhm THEN
        fMaxKOhm := fNegKOhm;                      // 负极更大 / the negative pole is larger
    END_IF
    fMinKOhm := fPosKOhm;                          // 极小值种子 / minimum seed
    IF fNegKOhm < fMinKOhm THEN
        fMinKOhm := fNegKOhm;                      // 负极更小 / the negative pole is smaller
    END_IF
    IF fMinKOhm > DL_SGF_TOL THEN
        fRatio := fMaxKOhm / fMinKOhm;             // 失衡比值（除子已判非零）[无量纲] / imbalance ratio
    ELSE
        fRatio := 1.0;                             // 极小值为零：比值不可算，按不失衡处理（不可判支路已前置）/ ratio unusable, treated as balanced
    END_IF
    bUnbalanced := (fRatio > DL_SGF_IMB_RATIO);    // 失衡判据 / imbalance predicate

    (*--------------------------------------------------------------------------
     * 段 9｜两级阈值确认与锁存：连续 nConfirmEff 拍低于阈值才置位，置位后锁存
     *       退化分支（绝缘哨兵）天然远高于阈值，不会触发，无需特判
     *-------------------------------------------------------------------------*)
    bAlarmNow := (fTotalKOhm < fAlarmKOhm);        // 告警判据 [kΩ] / alarm predicate
    bWarnNow := (fTotalKOhm < fWarnKOhm);          // 预警判据 [kΩ] / warning predicate
    IF bAlarmNow THEN
        IF nAlarmCnt < nConfirmEff THEN
            nAlarmCnt := nAlarmCnt + 1;            // 告警确认计数自增（上限即确认拍数）/ alarm counter increments up to the confirmation count
        END_IF
    ELSE
        nAlarmCnt := 0;                            // 断链即清零（防间歇性漏电被"攒"成告警）/ counter cleared on any drop-out
    END_IF
    IF bWarnNow THEN
        IF nWarnCnt < nConfirmEff THEN
            nWarnCnt := nWarnCnt + 1;              // 预警确认计数自增 / warning counter increments
        END_IF
    ELSE
        nWarnCnt := 0;                             // 断链即清零 / counter cleared
    END_IF
    IF nAlarmCnt >= nConfirmEff THEN
        bAlarm := TRUE;                            // 告警锁存（仅 bReset 可清）/ alarm latched, clearable only by reset
    END_IF
    IF nWarnCnt >= nConfirmEff THEN
        bWarn := TRUE;                             // 预警锁存（仅 bReset 可清）/ warning latched
    END_IF
    IF bAlarm THEN
        bWarn := TRUE;                             // 告警成立必然伴随预警（分级语义自洽）/ an alarm implies the warning
    END_IF

    (*--------------------------------------------------------------------------
     * 段 10｜出口码优先级：告警 > 预警 > 失衡提示 > 无错（同拍只能出一个码）
     *-------------------------------------------------------------------------*)
    IF bAlarm THEN
        eErr := 16#0000_0000;                      // 告警为状态量（bAlarm 出口），不占信息码位 / the alarm is a status, no info slot used
        eState := E_DL_StringInsState.eAlarm;      // 进告警监视相 / enter the alarm-monitoring state
    ELSIF bWarn THEN
        eErr := 16#0000_0000;                      // 预警同为状态量 / the warning is a status too
        eState := E_DL_StringInsState.eMeasure;    // 阻值仍有效，留在推算相 / resistances valid, stay in the measurement state
    ELSIF bUnbalanced THEN
        eErr := DL_SGF_CODE_INFO_2;                // 信息级：单极对地阻抗失衡提示 / info: single-pole imbalance hint
        eState := E_DL_StringInsState.eMeasure;    // 留推算相 / stay in the measurement state
    ELSE
        eErr := 16#0000_0000;                      // 无提示 / no hint
        eState := E_DL_StringInsState.eMeasure;    // 推算相 / measurement state
    END_IF
    IF bDegenerate AND (NOT bAlarm) AND (NOT bWarn) THEN
        eErr := 16#0000_0000;                      // 完全平衡（绝缘哨兵）无错，HMI 以饱和值显示 / balanced insulation reports no code
    END_IF
END_IF

(*------------------------------------------------------------------------------
 * 段 11｜状态机：CASE 含 ELSE 兜底（非法状态 → 035C + 阻值回零 + 许可撤）
 *       失能闸在此收口：不判、bValid := FALSE，但绝不清除已锁存的告警
 *----------------------------------------------------------------------------*)
CASE eState OF

    E_DL_StringInsState.eIdle:
        bValid := FALSE;                           // 失能闸显式不可用（R72）/ explicit FALSE on the disable gate
        fInsPosKOhm := DL_SGF_ZERO;                // 正极阻值回零 / positive resistance zeroed
        fInsNegKOhm := DL_SGF_ZERO;                // 负极阻值回零 / negative resistance zeroed
        fInsTotalKOhm := DL_SGF_ZERO;              // 并联阻值回零 / parallel resistance zeroed
        bUnbalanced := FALSE;                      // 失能不判失衡 / no imbalance verdict when disabled
        bUndecidable := FALSE;                     // 失能不报不可判 / no undecidable flag when disabled
        eErr := 16#0000_0000;                      // 待机无错 / no error in idle
        bError := FALSE;                           // 待机无故障 / no fault in idle
        // 失能绝不清除已锁存的 bWarn/bAlarm（历史事实，仅人工复位可清）/ a latched alarm survives a disable
        IF bEnable THEN
            eState := E_DL_StringInsState.eMeasure; // 使能进推算相 / enable enters the measurement state
            bFirstScan := FALSE;                   // 首拍标志清除 / first-scan flag cleared
        END_IF

    E_DL_StringInsState.eMeasure:
        bValid := TRUE;                            // 阻值可用 / resistances usable
        bError := FALSE;                           // 推算相无故障 / no fault on the measurement path
        IF NOT bEnable THEN
            eState := E_DL_StringInsState.eIdle;   // 失能回待机（退出条件一）/ disable, first exit
            bValid := FALSE;                       // 失能闸显式不可用 / explicit FALSE on the disable gate
        ELSIF bUndecidableNow THEN
            eState := E_DL_StringInsState.eUndecidable;   // 电压条件不成立转不可判（退出条件二）/ voltage conditions fail, second exit
        END_IF

    E_DL_StringInsState.eUndecidable:
        bValid := FALSE;                           // 阻值不可用（禁伪阻值，R42 家族）/ resistances unusable
        bError := FALSE;                           // 信息级不置 bError / info never raises bError
        eErr := DL_SGF_CODE_INFO_1;                // 信息级：绝缘推算不可判 / info: insulation not decidable
        IF NOT bEnable THEN
            eState := E_DL_StringInsState.eIdle;   // 失能回待机（退出条件一）/ disable, first exit
        ELSIF (NOT bUndecidableNow) THEN
            eState := E_DL_StringInsState.eMeasure;   // 电压条件恢复回推算相（退出条件二）/ conditions recovered, second exit
        END_IF

    E_DL_StringInsState.eAlarm:
        bValid := TRUE;                            // 阻值可用（告警期间继续监视）/ resistances usable, monitoring continues
        bError := FALSE;                           // 告警是状态量不是故障码 / an alarm is a status, not a fault code
        eErr := 16#0000_0000;                      // 不占信息码位 / no info slot used
        IF NOT bEnable THEN
            eState := E_DL_StringInsState.eIdle;   // 失能回待机（退出条件一，锁存保留）/ disable, first exit, the latch survives
            bValid := FALSE;                       // 失能闸显式不可用 / explicit FALSE on the disable gate
        ELSIF bUndecidableNow THEN
            eState := E_DL_StringInsState.eUndecidable;   // 电压条件不成立转不可判（退出条件二）/ undecidable, second exit
        ELSIF (NOT bAlarm) THEN
            eState := E_DL_StringInsState.eMeasure; // 复位清锁存后回推算相（退出条件三）/ latch cleared by reset, third exit
        END_IF

    E_DL_StringInsState.eFault:
        bValid := FALSE;                           // 故障闸显式不可用（R72）/ explicit FALSE on the fault gate
        bError := TRUE;                            // 故障级必置 bError（R45 配对）/ fault-class pairs with bError
        fInsPosKOhm := DL_SGF_ZERO;                // 正极阻值回零安全侧 / positive resistance zeroed, safe side
        fInsNegKOhm := DL_SGF_ZERO;                // 负极阻值回零安全侧 / negative resistance zeroed, safe side
        fInsTotalKOhm := DL_SGF_ZERO;              // 并联阻值回零安全侧 / parallel resistance zeroed, safe side
        bUnbalanced := FALSE;                      // 故障态不判失衡 / no imbalance verdict in fault
        bUndecidable := FALSE;                     // 故障态不报不可判 / no undecidable flag in fault
        IF eErr = 16#0000_0000 THEN
            eErr := DL_SGF_CODE_FLT_3;             // 入口无码时按非法状态兜底（R45：bError 必须有对应码）/ illegal-state fallback
        END_IF
        IF bEnable AND (fBridgeKOhm > DL_SGF_TOL) AND (fAlarmKOhm < fWarnKOhm - DL_SGF_TOL) THEN
            eState := E_DL_StringInsState.eIdle;   // 组态恢复且使能才回待机（退出条件 ≥2）/ recover only when the configuration is sane
        END_IF

    ELSE
        eState := E_DL_StringInsState.eFault;      // 非法状态兜底 / illegal-state fallback
        eErr := DL_SGF_CODE_FLT_3;                 // 故障级兜底：非法状态 / fault fallback: illegal state
        bError := TRUE;                            // 故障级必置 bError（R45 配对）/ fault-class pairs with bError
        bValid := FALSE;                           // 阻值不可用 / resistances unusable
        fInsPosKOhm := DL_SGF_ZERO;                // 正极阻值回零安全侧 / positive resistance zeroed, safe side
        fInsNegKOhm := DL_SGF_ZERO;                // 负极阻值回零安全侧 / negative resistance zeroed, safe side
        fInsTotalKOhm := DL_SGF_ZERO;              // 并联阻值回零安全侧 / parallel resistance zeroed, safe side
        bUnbalanced := FALSE;                      // 失衡标志撤 / imbalance withdrawn

END_CASE
END_FUNCTION_BLOCK

(* ---- FB_DL_UnscramblerSeq.st ---- *)
(*
  ==================================================================
  组件名 Component  : FB_DL_UnscramblerSeq
  分类   Category   : DL_Process
  前缀   Naming     : FB_DL_ ｜ b/n/u/f/t/e/st 类型前缀制（R265）
  码位   Code ID    : 16#0006_3038（故障级：卡瓶监视窗超时）｜ 16#0006_3039
                      （故障级：组态非法）
  版本   Version    : 1.0.1
  变更   CHANGELOG  : v1.0.1 _bHold 跨相粘滞统一清零
  复杂度 Complexity  : 中
  功能   Purpose    : 理瓶整理顺控：进瓶整理 → 乱瓶分拣 → 整理完成的相序推进，
                      卡瓶监视窗（卡瓶检测电平持续超窗即锁存故障）+ 料满停进
                      （满仓强制停进不 faults）；供理瓶机 / 提升料仓类工位。
  开源溯源 Origin    : OMAC PackML 状态模型（公开标准，T2-7 次源）：仅借 17 态
                      模型的相语义聚合口径（本件聚合为四相，R264 唯一声明）；
                      理瓶顺控逻辑完全自研，零代码复制。
  许可证 License    : MIT
  参考   Reference  : IEC 61131-3:2013 §6.6 状态机 / TON / R_TRIG 语义；
                      OMAC PackML 状态模型公开条款（借相语义，不抄文）
  平台   Platform   : 纯 IEC 61131-3（TON / R_TRIG / ENUM+CASE / 四则），三平台通用
  依赖   Depends    : 仅 Standard.library（TON / R_TRIG 属标准件）
  分工声明 Split     : FB_DL_CapSorterSeq（ caps 分拣专用顺控）/ FB_DL_FeederLevel
                      （料位控制）与本件互引；本件为理瓶相序 + 卡瓶保护 +
                      料满停进三合一工站级顺控，单相控制归各自属主（R216）。
  归属 Ownership     : E_DL_UnscrPhase 属主为本文件（全库唯一定义，R264）；
                      引用件只引用不重声明。
  ------------------------------------------------------------------
  边界 Boundary     :
                      一 组态闸结构早退（族② 判据，逐项点名 R272）：
                         tJamWin ≤ 0（卡瓶窗非正）或 tPhaseMin ≤ 0（相最短
                         驻留非正）→ 组态码 3039 + 三件套 + RETURN；
                      二 状态机 ENUM + CASE 必带 ELSE（非法态兜底落 eFault +
                         锁存 3039，禁静默）；本拍合法事件（停止 / 料满 /
                         相完成沿）优先于卡瓶超时迁移（R275 同拍竞态）；
                      三 卡瓶窗口径：bJamSense 电平 + tJamWin 持续超窗 →
                         锁存 3038；瞬时卡瓶抖动由窗吸收（窗时长须大于
                         检测去抖上限，交付默认 T#3S，调用方改参须维持）；
                      四 失败锁存 bJamFault + _bFaultLatch；锁存解除式
                         （可达自证，R152）：bResetCmd 上升沿清锁存回 eIdle
                         （输入引脚恒可达，无「置位即永久」路径）；
                      五 料满停进语义（不 faults）：bHopperFull 电平在
                         eFeed / eSort 相强制 bFeedOut = FALSE 停进、相保持
                         挂起（相驻留最短时限 tonPhase 在料满期同步挂起，
                         防满仓期被误判相超时——挂相不挂故障）；料满解除
                         后相序自动续推；
                      六 bEnable = FALSE 的语义写死（FB33-4 声明行）：强制
                         eIdle + 双出口复位（不 faults，使能断开 ≠ 顺控故障）；
                      七 TON / R_TRIG 段 0 无条件刷新（禁入分支，R7）；监视
                         TON IN 串故障锁存门控（FB50-1）；相驻留 TON 为
                         「最短驻留门槛」口径（IN 串相条件，到时即允许
                         迁移，不是超时故障源）；
                      八 首拍 _bInit 全量初始化；无浮点量、无除法；无全局、
                         无外部变量、无物理地址。
  错误码 Codes      :
    16#0006_3038【故障级】卡瓶持续超窗（bJamSense 持续 tJamWin，疑似卡瓶 /
                         检测回路故障）
    16#0006_3039【故障级】组态非法（tJamWin ≤ 0 / tPhaseMin ≤ 0）或非法状态
                         拦截（ELSE 兜底）
  码位反证 Note     :
    3038 与 3039 不可合并：3038 与组态无关（需运行期卡瓶电平到达，处置人 =
    现场机务），3039 组态即刻判（处置人 = 组态工程师），可由场景还原（R90），
    分立；料满停进不设码（停进不是故障，边界五语义声明）。
  验收 Acceptance   :
    算法已证（脚本）：未跑 ｜ 编译器已证（三平台）：未跑
    V1 启动 → eFeed（bFeedOut = TRUE）；相驻留到时 + 分拣使能 → eSort
    V2 分拣完成信号 → eReady（bFeedOut / bSortOut 复位）
    V3 bJamSense 持续超窗 → 锁存 3038、双出口切断
    V4 瞬时卡瓶 < 窗 → 不误报（窗吸收向量）
    V5 eFeed 期料满 → bFeedOut 强制 FALSE、相挂起不超时（边界五向量）
    V6 tJamWin = T#0S → 组态早退 3039；V7 失能 → eIdle 双出口复位
    V8 非法枚举态（强改 eState）→ ELSE 兜底落 eFault + 3039
  修订记录 Revision  :
    2026-11-21  v1.0.0  R64 首版（批 3 · 序号 10，PackML 相语义 + 自研顺控）
    2026-11-22  v1.0.1  R65 点修（_bHold 跨相粘滞，R64 终审项）：v1.0.0 中
                        _bHold 仅在 eFeed / eSort 相内随料满电平置清，迁移
                        出口（停止回 eIdle / 分拣完成迁 eReady / 锁存落
                        eFault）不清 _bHold，跨相粘滞使下一拍 tonPhase
                        （串 NOT _bHold 门控）在非保持相读到旧值；v1.0.1
                        采用统一入口清零式（择一实现声明）：在段 0 顶部
                        （定时器刷新之前，保证同拍收敛）对非保持相强制
                        _bHold := FALSE，理由——迁移出口分散于两相共 5 处，
                        逐出口补清易漏且新增出口须重复纪律，单点集中清零
                        全覆盖；eFeed / eSort 相内料满置清语义不受影响
  ==================================================================
*)
TYPE E_DL_UnscrPhase :
(
    eIdle  := 0,  // 待机：等启动 / idle, waiting for the start
    eFeed  := 10, // 进瓶整理：进料出口有效，等相驻留 / the feed phase with the feed outlet
    eSort  := 20, // 乱瓶分拣：分拣出口有效，等完成信号 / the sort phase with the sort outlet
    eReady := 30, // 整理完成：双出口复位，等再启动或停止 / the ready phase with both outlets reset
    eFault := 40  // 锁存故障：卡瓶超窗或非法态，复位沿解除 / a latched fault released by the reset edge
);
END_TYPE

FUNCTION_BLOCK FB_DL_UnscramblerSeq
VAR_INPUT
    bEnable    : BOOL := TRUE;   // 使能，FALSE 时强制 eIdle + 双出口复位（边界六）/ the enable, false forces the idle and resets both outlets
    bStart     : BOOL := FALSE;  // 启动电平 [-]（eReady / eIdle 相生效）/ the start level valid in the ready and idle phases
    bSortEn    : BOOL := FALSE;  // 分拣使能电平 [-]（eFeed → eSort 的迁移前提）/ the sort enable as the transition premise
    bSortDone  : BOOL := FALSE;  // 分拣完成电平 [-]（eSort → eReady 的事件）/ the sort done event of the sort phase
    bJamSense  : BOOL := FALSE;  // 卡瓶检测电平 [-] / the jam detection level
    bHopperFull: BOOL := FALSE;  // 料满电平 [-]（满仓停进，不 faults，边界五）/ the hopper full level stopping the feed without a fault
    bResetCmd  : BOOL := FALSE;  // 故障复位电平，上升沿清锁存回 eIdle（边界四解除式）/ the fault reset level, its rising edge releases the latch
    tJamWin    : TIME := T#3S;   // 卡瓶监视窗 [毫秒]，须 > 0 / the jam window, positive
    tPhaseMin  : TIME := T#2S;   // 相最短驻留 [毫秒]，须 > 0 / the minimum phase dwell, positive
END_VAR
VAR_OUTPUT
    bFeedOut : BOOL := FALSE;           // 进料出口 [-]（料满 / 故障 / 失能强制 FALSE）/ the feed outlet forced false on full, fault or disable
    bSortOut : BOOL := FALSE;           // 分拣出口 [-]（故障 / 失能强制 FALSE）/ the sort outlet forced false on a fault or disable
    bJamFault: BOOL := FALSE;           // 卡瓶故障（锁存）[-] / the latched jam fault
    eState   : E_DL_UnscrPhase;         // 状态机出口 [状态] / the state machine outlet
    bValid   : BOOL := FALSE;           // 判据可用 [-] / the criteria are usable
    eErr     : UDINT := 16#0000_0000;   // 错误码，0 = 正常 / the error code, zero is ok
    bError   : BOOL := FALSE;           // 故障标志（故障级码同拍置位，R45 配对）/ the fault flag raised with a fault level code
END_VAR
VAR
    _bInit      : BOOL := FALSE;  // 首拍初始化标志（R310 / FB50-2）/ the first scan flag
    _eState     : E_DL_UnscrPhase := E_DL_UnscrPhase.eIdle; // 内部状态寄存器 / the internal state register
    _bFaultLatch: BOOL := FALSE;  // 故障锁存副本（仅复位沿清除）/ the fault latch copy
    _uLatch     : UDINT := 16#0000_0000; // 故障码锁存 [码]（复位沿清除，FB33-1）/ the latched fault code cleared by the reset edge
    _bCfgBad    : BOOL := FALSE;  // 组态非法标记（逐拍重算）/ the configuration fault flag
    _bHold      : BOOL := FALSE;  // 料满挂相标记（料满期相驻留计时同步挂起，边界五）/ the hold flag suspending the dwell timer on full
    rtReset     : R_TRIG;         // 复位沿实例，段 0 无条件刷新（R7）/ the reset edge instance refreshed unconditionally
    tonJam      : TON;            // 卡瓶监视窗定时器，段 0 无条件刷新 / the jam window timer refreshed unconditionally
    tonPhase    : TON;            // 相最短驻留定时器（最短驻留门槛口径，边界七）/ the phase dwell floor timer
END_VAR  // R64 结构补齐：VAR 段缺失的 END_VAR（门禁机械修复）
VAR CONSTANT
    DL_UNP_TIME0 : TIME := T#0S;          // 时间零常量 [毫秒] / the time zero constant
    DL_UNP_ZEROU : UDINT := 16#0000_0000; // 码零常量 / the code zero constant
END_VAR

// 段 0a｜_bHold 跨相粘滞统一清零（v1.0.1，R64 终审项修复；置段 0 之前保证
//         tonPhase 同拍读到新值）/ segment 0a, the unified sticky clear of the hold flag
IF (_eState <> E_DL_UnscrPhase.eFeed) AND (_eState <> E_DL_UnscrPhase.eSort) THEN // 非保持相（eIdle / eReady / eFault）/ outside the holding phases
    _bHold := FALSE; // 非保持相强制清挂相标记（防跨相粘滞；eFeed / eSort 相内料满置清语义不受影响，v1.0.1 择统一式理由见修订记录）/ clear the hold flag outside the holding phases
END_IF

// 段 0｜定时器与沿检测无条件周期刷新（禁入分支，R7；监视 TON 串锁存门控，FB50-1）/ segment 0, the unconditional refresh
rtReset(CLK := bResetCmd); // 复位沿 / the reset edge
tonJam(IN := (( _eState = E_DL_UnscrPhase.eFeed) OR (_eState = E_DL_UnscrPhase.eSort))
          AND bJamSense AND (NOT _bFaultLatch), PT := tJamWin); // 卡瓶窗计时（仅进瓶 / 分拣相有效，串锁存门控防复位同拍重锁）/ the jam window only in the feed and sort phases with the latch gate
tonPhase(IN := (( _eState = E_DL_UnscrPhase.eFeed) OR (_eState = E_DL_UnscrPhase.eSort))
          AND (NOT _bHold) AND (NOT _bFaultLatch), PT := tPhaseMin); // 相驻留计时（料满挂相机同步挂起，边界五；最短驻留门槛口径，边界七）/ the dwell timer suspended on the hold, a floor not a timeout source

// 段 1｜首拍初始化与复位沿作用域（R310 / R311）/ segment 1, the first scan init and the reset edge scope
IF NOT _bInit THEN // 首拍一拍 / the first scan
    _bInit := TRUE; // 置首拍标志 / raise the first scan flag
    _eState := E_DL_UnscrPhase.eIdle; // 状态显式落空闲 / place the state to idle
    _bFaultLatch := FALSE; // 故障锁存显式清零 / clear the fault latch explicitly
    _uLatch := DL_UNP_ZEROU; // 码锁存显式清零 / clear the latched code explicitly
    _bHold := FALSE; // 挂相标记显式清零 / clear the hold flag explicitly
END_IF
IF rtReset.Q THEN // 复位沿（作用域声明：清锁存 + 迁相位 + 清挂相，R311）/ the reset edge with the declared scope
    _bFaultLatch := FALSE; // 清故障锁存（唯一解除路径，边界四自证可达）/ clear the fault latch, the only release path
    _uLatch := DL_UNP_ZEROU; // 清码锁存 / clear the latched code
    _eState := E_DL_UnscrPhase.eIdle; // 迁回空闲 / back to idle
    _bHold := FALSE; // 清挂相标记 / clear the hold flag
END_IF

// 段 2｜组态域闸结构早退（边界一，族② 判据：两时限逐项点名）/ segment 2, the structural early exit on an illegal configuration
_bCfgBad := (tJamWin <= DL_UNP_TIME0) OR (tPhaseMin <= DL_UNP_TIME0); // 组态非法（任一窗非正）/ an illegal configuration
IF _bCfgBad THEN // 组态非法：结构早退（出口三件套 + RETURN）/ an illegal configuration exits structurally
    eState := _eState; // 状态照实出口（冻结）/ export the state as is
    bFeedOut := FALSE; // 进料出口切断（组态非法期禁下发）/ cut the feed outlet off
    bSortOut := FALSE; // 分拣出口切断 / cut the sort outlet off
    bJamFault := _bFaultLatch; // 故障锁存照实回放 / replay the latch
    bValid := FALSE; // 判据不可用 / the criteria are not usable
    eErr := 16#0006_3039; // 故障级：组态非法 / fault grade, an illegal configuration
    bError := TRUE; // 同拍置故障标志（R45 配对）/ raise the fault flag on the same scan
    RETURN; // 结构早退 / the structural early exit
END_IF

// 段 3｜失能分支：强制 eIdle + 双出口复位，不 faults（边界六声明行）/ segment 3, the disabled branch
IF NOT bEnable THEN // 失能 / disabled
    _eState := E_DL_UnscrPhase.eIdle; // 强制空闲 / force the idle
    _bFaultLatch := FALSE; // 锁存复位（使能断开 ≠ 顺控故障）/ clear the latch
    _uLatch := DL_UNP_ZEROU; // 码锁存复位 / clear the code
    _bHold := FALSE; // 挂相标记复位 / clear the hold flag
    eState := _eState; // 状态出口 / the state outlet
    bFeedOut := FALSE; // 进料出口复位 / the feed outlet resets
    bSortOut := FALSE; // 分拣出口复位 / the sort outlet resets
    bJamFault := FALSE; // 故障位复位 / the fault bit resets
    bValid := FALSE; // 失能即不可用 / the criteria are not usable while disabled
    bError := FALSE; // 失能不是故障 / a disabled device is not a fault
    eErr := DL_UNP_ZEROU; // 失能不发码 / no code is emitted while disabled
    RETURN; // 早退 / early return
END_IF

// 段 4｜主状态机（ENUM + CASE，ELSE 兜底；本拍合法事件优先于卡瓶超时，R275）/ segment 4, the main machine, the legal event before the jam timeout
CASE _eState OF
    E_DL_UnscrPhase.eIdle: // 空闲相 / the idle phase
        IF bStart AND (NOT _bFaultLatch) AND (NOT _bCfgBad) THEN // 启动电平 + 全量闸位复检（R274）/ the start with the full gate recheck
            _eState := E_DL_UnscrPhase.eFeed; // 迁入进瓶相 / enter the feed phase
        END_IF
    E_DL_UnscrPhase.eFeed: // 进瓶相（本拍合法事件优先：停止 / 分拣使能迁移先消化，再消化卡瓶超窗，R275）/ the feed phase, the legal event before the jam timeout
        IF bHopperFull THEN // 料满停进：相挂起不迁相（边界五，挂相不挂故障）/ the full level holds the phase without a fault
            _bHold := TRUE; // 置挂相标记（tonPhase 同步挂起，防满仓误判）/ raise the hold flag
        ELSE // 料满解除 / the full level released
            _bHold := FALSE; // 清挂相标记（相序自动续推）/ clear the hold flag
        END_IF
        IF NOT bStart THEN // 事件优先：停止电平 / the stop level, the event goes first
            _eState := E_DL_UnscrPhase.eIdle; // 回空闲 / back to idle
        ELSIF tonPhase.Q AND bSortEn THEN // 相驻留到时 + 分拣使能（迁移门槛齐备）/ the dwell floor reached with the sort enable
            _eState := E_DL_UnscrPhase.eSort; // 迁入分拣相 / enter the sort phase
        ELSIF tonJam.Q THEN // 卡瓶持续超窗（卡瓶判据，真实可达：瓶体楔死）/ the jam stayed through the window, reachable by a wedged bottle
            _bFaultLatch := TRUE; // 锁存故障 / latch the fault
            _uLatch := 16#0006_3038; // 故障级：卡瓶超窗 / fault grade, the jam through the window
            bError := TRUE; // 同拍置故障标志（R45 配对，段 6 故障分支沿用）/ raise the fault flag on the same scan
        END_IF
    E_DL_UnscrPhase.eSort: // 分拣相（同拍序与 eFeed 一致，R275）/ the sort phase with the same event order
        IF bHopperFull THEN // 料满挂相（分拣出口保持，进料出口停，边界五）/ the full level holds the phase, the sort outlet stays
            _bHold := TRUE; // 置挂相标记 / raise the hold flag
        ELSE // 料满解除 / the full level released
            _bHold := FALSE; // 清挂相标记 / clear the hold flag
        END_IF
        IF NOT bStart THEN // 事件优先：停止电平 / the stop level, the event goes first
            _eState := E_DL_UnscrPhase.eIdle; // 回空闲 / back to idle
        ELSIF bSortDone THEN // 事件优先：分拣完成 / the sort done, the event goes first
            _eState := E_DL_UnscrPhase.eReady; // 迁入完成相 / enter the ready phase
        ELSIF tonJam.Q THEN // 卡瓶持续超窗 / the jam through the window
            _bFaultLatch := TRUE; // 锁存故障 / latch the fault
            _uLatch := 16#0006_3038; // 故障级：卡瓶超窗 / fault grade, the jam through the window
            bError := TRUE; // 同拍置故障标志（R45 配对，段 6 故障分支沿用）/ raise the fault flag on the same scan
        END_IF
    E_DL_UnscrPhase.eReady: // 完成相（整理完成驻留，等再启动或停止）/ the ready phase dwelling for the next start or stop
        IF NOT bStart THEN // 停止电平 / the stop level
            _eState := E_DL_UnscrPhase.eIdle; // 回空闲 / back to idle
        ELSIF bStart AND (NOT bHopperFull) THEN // 再启动且料已不满（料满期不重进，防顶仓）/ a restart with the hopper not full
            _eState := E_DL_UnscrPhase.eFeed; // 重进进瓶相 / reenter the feed phase
        END_IF
    E_DL_UnscrPhase.eFault: // 锁存故障相（驻留，解除由段 1 复位沿承担）/ the fault phase dwelling, the release belongs to the reset edge
        ; // 驻留语义由注释表达（禁自赋值死语句，R261）/ the dwell is expressed by this comment without a dead statement
    ELSE // 非法枚举值拦截（边界二：落故障相并锁存，禁静默）/ the illegal enumeration guard
        _bFaultLatch := TRUE; // 锁存故障 / latch the fault
        _uLatch := 16#0006_3039; // 故障级：非法状态拦截（归入组态族一码，出口同形，R90）/ fault grade, the illegal state in the configuration family
        bError := TRUE; // 同拍置故障标志（R45 配对）/ raise the fault flag on the same scan
        _eState := E_DL_UnscrPhase.eFault; // 落故障相 / force the fault phase
END_CASE

// 段 5｜故障锁存迁移闸（置于解除段之后防同拍抢迁，R258）/ segment 5, the latch to phase gate
IF _bFaultLatch AND (_eState <> E_DL_UnscrPhase.eFault) THEN // 已锁存但不在故障相 / latched outside the fault phase
    _eState := E_DL_UnscrPhase.eFault; // 迁入故障相 / enter the fault phase
END_IF

// 段 6｜统一出口（名实双出口同源，R191）/ segment 6, the unified outlet
eState := _eState; // 状态出口 / the state outlet
bFeedOut := (_eState = E_DL_UnscrPhase.eFeed) AND (NOT _bHold)
         AND (NOT _bFaultLatch); // 进料出口与状态 / 挂相 / 锁存同源派生（边界五料满停进）/ the feed outlet derived from the state, the hold and the latch
bSortOut := (_eState = E_DL_UnscrPhase.eSort) AND (NOT _bFaultLatch); // 分拣出口与状态 / 锁存同源派生（料满期分拣出口保持，边界五）/ the sort outlet derived from the state and the latch
bJamFault := _bFaultLatch; // 故障位与锁存同源 / the fault bit from the latch
bValid := (NOT _bFaultLatch) AND (NOT _bCfgBad); // 判据可用（无锁存且组态合法）/ usable without a latch and with a legal configuration
IF _bFaultLatch THEN // 故障锁存回放优先（不在故障相按当下输入重新推断，R152）/ the latched fault replays first
    bValid := FALSE; // 故障相不可用 / not usable in the fault phase
    bError := TRUE; // 故障位置位（R45 配对）/ raise the fault bit
    eErr := _uLatch; // 锁存码回放 / replay the latched code
ELSE // 无事件 / no event
    bError := FALSE; // 无故障 / no fault
    eErr := DL_UNP_ZEROU; // 正常 / ok
END_IF
END_FUNCTION_BLOCK
